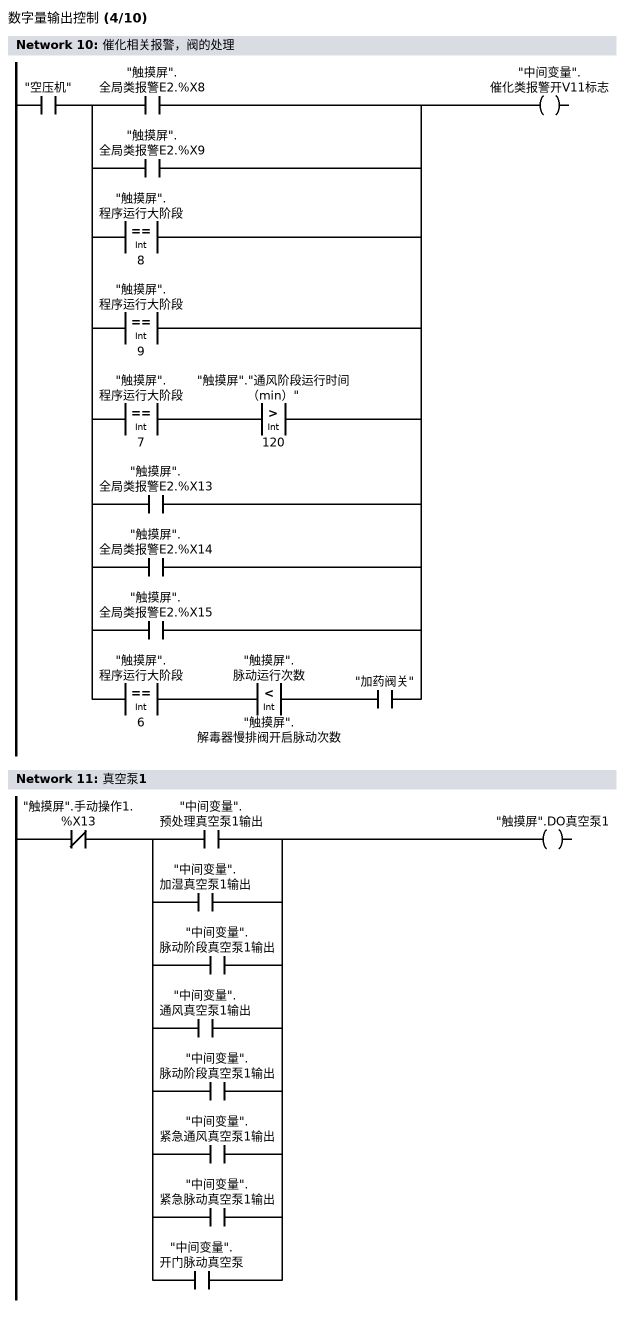
   RUNG wire#powerrail
      Contact( "空压机" )
      wire#w1
      Contact( "触摸屏".全局类报警E2.%X8 )
      wire#w2
      Coil( "中间变量".催化类报警开V11标志 )
   END_RUNG
   RUNG wire#w1
      Contact( "触摸屏".全局类报警E2.%X9 )
   END_RUNG wire#w2
   RUNG wire#w1
      { S7_Templates := "SrcType := Int" } EQ_Contact(in1 := "触摸屏".程序运行大阶段, in2 := 8)
   END_RUNG wire#w2
   RUNG wire#w1
      { S7_Templates := "SrcType := Int" } EQ_Contact(in1 := "触摸屏".程序运行大阶段, in2 := 9)
   END_RUNG wire#w2
   RUNG wire#w1
      { S7_Templates := "SrcType := Int" } EQ_Contact(in1 := "触摸屏".程序运行大阶段, in2 := 7)
      { S7_Templates := "SrcType := Int" } GT_Contact(in1 := "触摸屏"."通风阶段运行时间（min）", in2 := 120)
   END_RUNG wire#w2
   RUNG wire#w1
      Contact( "触摸屏".全局类报警E2.%X13 )
   END_RUNG wire#w2
   RUNG wire#w1
      Contact( "触摸屏".全局类报警E2.%X14 )
   END_RUNG wire#w2
   RUNG wire#w1
      Contact( "触摸屏".全局类报警E2.%X15 )
   END_RUNG wire#w2
   RUNG wire#w1
      { S7_Templates := "SrcType := Int" } EQ_Contact(in1 := "触摸屏".程序运行大阶段, in2 := 6)
      { S7_Templates := "SrcType := Int" } LT_Contact(in1 := "触摸屏".脉动运行次数, in2 := "触摸屏".解毒器慢排阀开启脉动次数)
      Contact( "加药阀关" )
   END_RUNG wire#w2
   // the same network as SCL:
   "中间变量".催化类报警开V11标志 := "空压机" AND ("触摸屏".全局类报警E2.%X8 OR "触摸屏".全局类报警E2.%X9 OR ("触摸屏".程序运行大阶段 = 8) OR ("触摸屏".程序运行大阶段 = 9) OR (("触摸屏".程序运行大阶段 = 7) AND ("触摸屏"."通风阶段运行时间（min）" > 120)) OR "触摸屏".全局类报警E2.%X13 OR "触摸屏".全局类报警E2.%X14 OR "触摸屏".全局类报警E2.%X15 OR (("触摸屏".程序运行大阶段 = 6) AND ("触摸屏".脉动运行次数 < "触摸屏".解毒器慢排阀开启脉动次数) AND "加药阀关"));
END_REGION

REGION Network 11: 真空泵1
   RUNG wire#powerrail
      I_Contact( "触摸屏".手动操作1.%X13 )
      wire#w1
      Contact( "中间变量".预处理真空泵1输出 )
      wire#w2
      Coil( "触摸屏".DO真空泵1 )
   END_RUNG
   RUNG wire#w1
      Contact( "中间变量".加湿真空泵1输出 )
   END_RUNG wire#w2
   RUNG wire#w1
      Contact( "中间变量".脉动阶段真空泵1输出 )
   END_RUNG wire#w2
   RUNG wire#w1
      Contact( "中间变量".通风真空泵1输出 )
   END_RUNG wire#w2
   RUNG wire#w1
      Contact( "中间变量".脉动阶段真空泵1输出 )
   END_RUNG wire#w2
   RUNG wire#w1
      Contact( "中间变量".紧急通风真空泵1输出 )
   END_RUNG wire#w2
   RUNG wire#w1
      Contact( "中间变量".紧急脉动真空泵1输出 )
   END_RUNG wire#w2
   RUNG wire#w1
      Contact( "中间变量".开门脉动真空泵 )
   END_RUNG wire#w2
   // the same network as SCL:
   "触摸屏".DO真空泵1 := NOT "触摸屏".手动操作1.%X13 AND ("中间变量".预处理真空泵1输出 OR "中间变量".加湿真空泵1输出 OR "中间变量".脉动阶段真空泵1输出 OR "中间变量".通风真空泵1输出 OR "中间变量".脉动阶段真空泵1输出 OR "中间变量".紧急通风真空泵1输出 OR "中间变量".紧急脉动真空泵1输出 OR "中间变量".开门脉动真空泵);
END_REGION

REGION Network 12: 真空泵2
END_REGION

REGION Network 13: 空压机
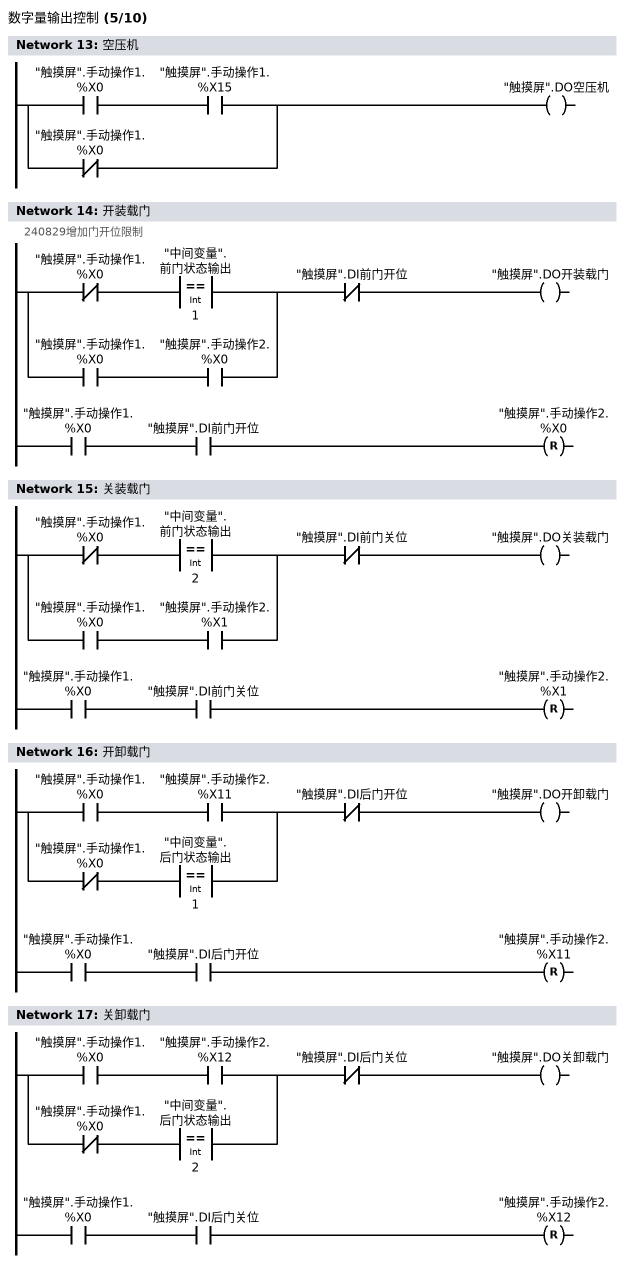
   RUNG wire#powerrail
      Contact( "触摸屏".手动操作1.%X0 )
      Contact( "触摸屏".手动操作1.%X15 )
      wire#w1
      Coil( "触摸屏".DO空压机 )
   END_RUNG
   RUNG wire#powerrail
      I_Contact( "触摸屏".手动操作1.%X0 )
   END_RUNG wire#w1
   // the same network as SCL:
   "触摸屏".DO空压机 := ("触摸屏".手动操作1.%X0 AND "触摸屏".手动操作1.%X15) OR NOT "触摸屏".手动操作1.%X0;
END_REGION

REGION Network 14: 开装载门
   // 240829增加门开位限制
   RUNG wire#powerrail
      I_Contact( "触摸屏".手动操作1.%X0 )
      { S7_Templates := "SrcType := Int" } EQ_Contact(in1 := "中间变量".前门状态输出, in2 := 1)
      wire#w1
      I_Contact( "触摸屏".DI前门开位 )
      Coil( "触摸屏".DO开装载门 )
   END_RUNG
   RUNG wire#powerrail
      Contact( "触摸屏".手动操作1.%X0 )
      Contact( "触摸屏".手动操作2.%X0 )
   END_RUNG wire#w1
   RUNG wire#powerrail
      Contact( "触摸屏".手动操作1.%X0 )
      Contact( "触摸屏".DI前门开位 )
      R_Coil( "触摸屏".手动操作2.%X0 )
   END_RUNG
   // the same network as SCL:
   "触摸屏".DO开装载门 := ((NOT "触摸屏".手动操作1.%X0 AND ("中间变量".前门状态输出 = 1)) OR ("触摸屏".手动操作1.%X0 AND "触摸屏".手动操作2.%X0)) AND NOT "触摸屏".DI前门开位;
   IF "触摸屏".手动操作1.%X0 AND "触摸屏".DI前门开位 THEN "触摸屏".手动操作2.%X0 := FALSE; END_IF;
END_REGION

REGION Network 15: 关装载门
   RUNG wire#powerrail
      I_Contact( "触摸屏".手动操作1.%X0 )
      { S7_Templates := "SrcType := Int" } EQ_Contact(in1 := "中间变量".前门状态输出, in2 := 2)
      wire#w1
      I_Contact( "触摸屏".DI前门关位 )
      Coil( "触摸屏".DO关装载门 )
   END_RUNG
   RUNG wire#powerrail
      Contact( "触摸屏".手动操作1.%X0 )
      Contact( "触摸屏".手动操作2.%X1 )
   END_RUNG wire#w1
   RUNG wire#powerrail
      Contact( "触摸屏".手动操作1.%X0 )
      Contact( "触摸屏".DI前门关位 )
      R_Coil( "触摸屏".手动操作2.%X1 )
   END_RUNG
   // the same network as SCL:
   "触摸屏".DO关装载门 := ((NOT "触摸屏".手动操作1.%X0 AND ("中间变量".前门状态输出 = 2)) OR ("触摸屏".手动操作1.%X0 AND "触摸屏".手动操作2.%X1)) AND NOT "触摸屏".DI前门关位;
   IF "触摸屏".手动操作1.%X0 AND "触摸屏".DI前门关位 THEN "触摸屏".手动操作2.%X1 := FALSE; END_IF;
END_REGION

REGION Network 16: 开卸载门
   RUNG wire#powerrail
      Contact( "触摸屏".手动操作1.%X0 )
      Contact( "触摸屏".手动操作2.%X11 )
      wire#w1
      I_Contact( "触摸屏".DI后门开位 )
      Coil( "触摸屏".DO开卸载门 )
   END_RUNG
   RUNG wire#powerrail
      I_Contact( "触摸屏".手动操作1.%X0 )
      { S7_Templates := "SrcType := Int" } EQ_Contact(in1 := "中间变量".后门状态输出, in2 := 1)
   END_RUNG wire#w1
   RUNG wire#powerrail
      Contact( "触摸屏".手动操作1.%X0 )
      Contact( "触摸屏".DI后门开位 )
      R_Coil( "触摸屏".手动操作2.%X11 )
   END_RUNG
   // the same network as SCL:
   "触摸屏".DO开卸载门 := (("触摸屏".手动操作1.%X0 AND "触摸屏".手动操作2.%X11) OR (NOT "触摸屏".手动操作1.%X0 AND ("中间变量".后门状态输出 = 1))) AND NOT "触摸屏".DI后门开位;
   IF "触摸屏".手动操作1.%X0 AND "触摸屏".DI后门开位 THEN "触摸屏".手动操作2.%X11 := FALSE; END_IF;
END_REGION

REGION Network 17: 关卸载门
   RUNG wire#powerrail
      Contact( "触摸屏".手动操作1.%X0 )
      Contact( "触摸屏".手动操作2.%X12 )
      wire#w1
      I_Contact( "触摸屏".DI后门关位 )
      Coil( "触摸屏".DO关卸载门 )
   END_RUNG
   RUNG wire#powerrail
      I_Contact( "触摸屏".手动操作1.%X0 )
      { S7_Templates := "SrcType := Int" } EQ_Contact(in1 := "中间变量".后门状态输出, in2 := 2)
   END_RUNG wire#w1
   RUNG wire#powerrail
      Contact( "触摸屏".手动操作1.%X0 )
      Contact( "触摸屏".DI后门关位 )
      R_Coil( "触摸屏".手动操作2.%X12 )
   END_RUNG
   // the same network as SCL:
   "触摸屏".DO关卸载门 := (("触摸屏".手动操作1.%X0 AND "触摸屏".手动操作2.%X12) OR (NOT "触摸屏".手动操作1.%X0 AND ("中间变量".后门状态输出 = 2))) AND NOT "触摸屏".DI后门关位;
   IF "触摸屏".手动操作1.%X0 AND "触摸屏".DI后门关位 THEN "触摸屏".手动操作2.%X12 := FALSE; END_IF;
END_REGION

REGION Network 18: 蜂鸣器FM
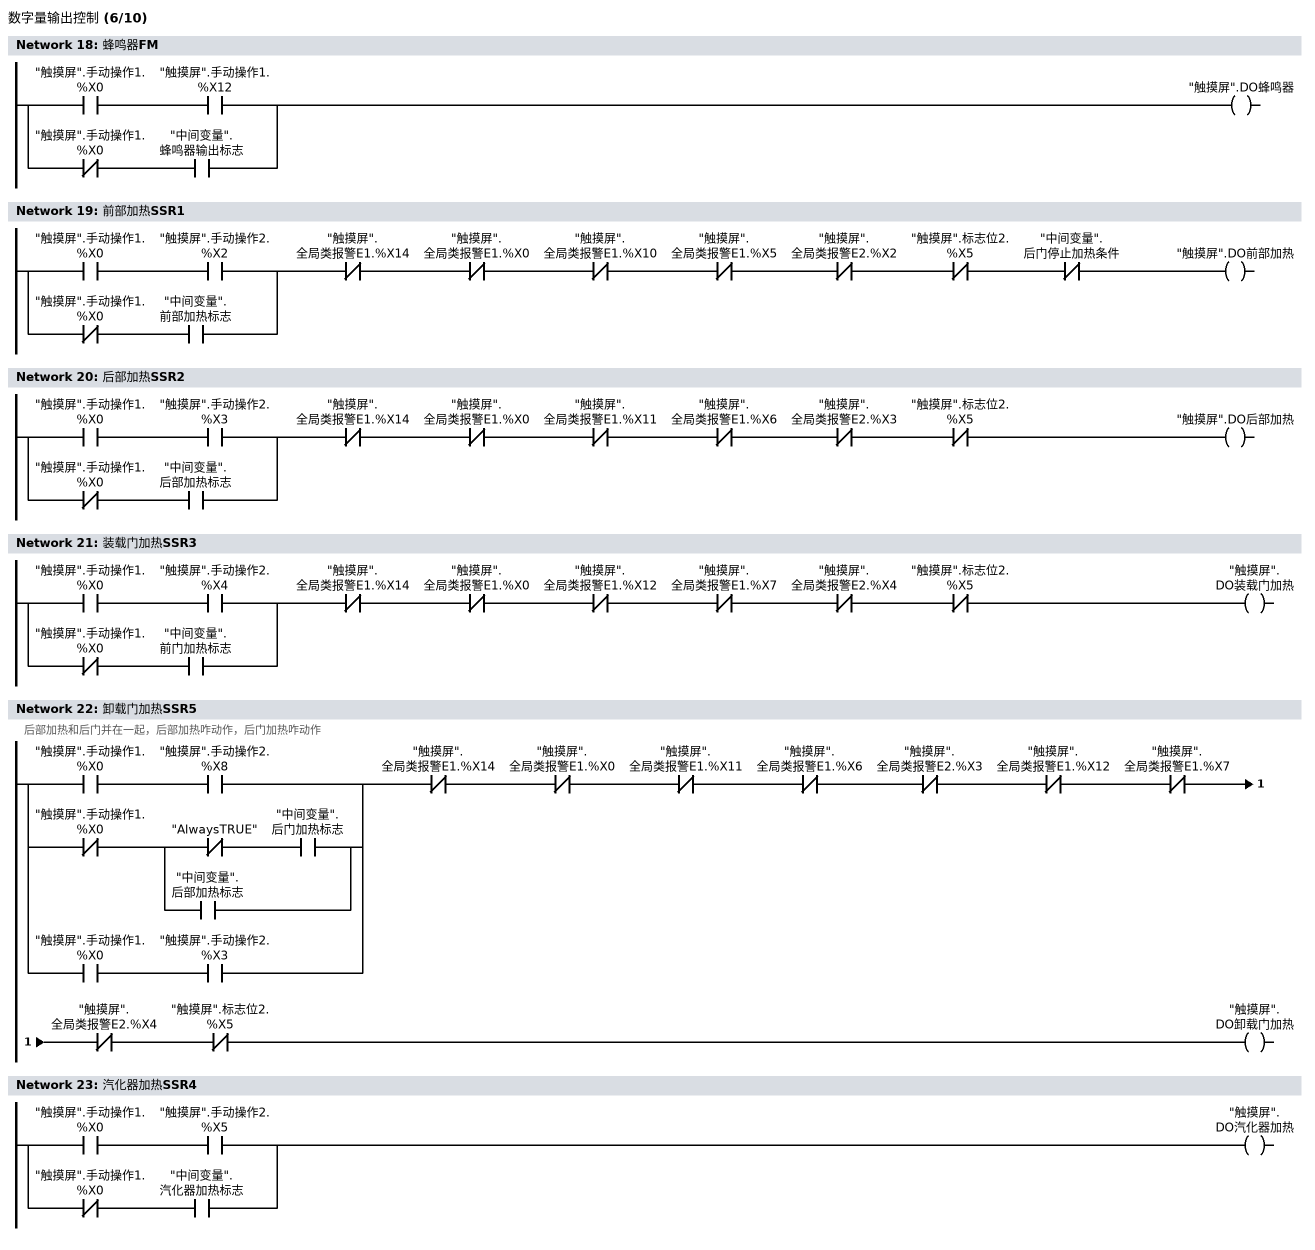
   RUNG wire#powerrail
      Contact( "触摸屏".手动操作1.%X0 )
      Contact( "触摸屏".手动操作1.%X12 )
      wire#w1
      Coil( "触摸屏".DO蜂鸣器 )
   END_RUNG
   RUNG wire#powerrail
      I_Contact( "触摸屏".手动操作1.%X0 )
      Contact( "中间变量".蜂鸣器输出标志 )
   END_RUNG wire#w1
   // the same network as SCL:
   "触摸屏".DO蜂鸣器 := ("触摸屏".手动操作1.%X0 AND "触摸屏".手动操作1.%X12) OR (NOT "触摸屏".手动操作1.%X0 AND "中间变量".蜂鸣器输出标志);
END_REGION

REGION Network 19: 前部加热SSR1
   RUNG wire#powerrail
      Contact( "触摸屏".手动操作1.%X0 )
      Contact( "触摸屏".手动操作2.%X2 )
      wire#w1
      I_Contact( "触摸屏".全局类报警E1.%X14 )
      I_Contact( "触摸屏".全局类报警E1.%X0 )
      I_Contact( "触摸屏".全局类报警E1.%X10 )
      I_Contact( "触摸屏".全局类报警E1.%X5 )
      I_Contact( "触摸屏".全局类报警E2.%X2 )
      I_Contact( "触摸屏".标志位2.%X5 )
      I_Contact( "中间变量".后门停止加热条件 )
      Coil( "触摸屏".DO前部加热 )
   END_RUNG
   RUNG wire#powerrail
      I_Contact( "触摸屏".手动操作1.%X0 )
      Contact( "中间变量".前部加热标志 )
   END_RUNG wire#w1
   // the same network as SCL:
   "触摸屏".DO前部加热 := (("触摸屏".手动操作1.%X0 AND "触摸屏".手动操作2.%X2) OR (NOT "触摸屏".手动操作1.%X0 AND "中间变量".前部加热标志)) AND NOT "触摸屏".全局类报警E1.%X14 AND NOT "触摸屏".全局类报警E1.%X0 AND NOT "触摸屏".全局类报警E1.%X10 AND NOT "触摸屏".全局类报警E1.%X5 AND NOT "触摸屏".全局类报警E2.%X2 AND NOT "触摸屏".标志位2.%X5 AND NOT "中间变量".后门停止加热条件;
END_REGION

REGION Network 20: 后部加热SSR2
   RUNG wire#powerrail
      Contact( "触摸屏".手动操作1.%X0 )
      Contact( "触摸屏".手动操作2.%X3 )
      wire#w1
      I_Contact( "触摸屏".全局类报警E1.%X14 )
      I_Contact( "触摸屏".全局类报警E1.%X0 )
      I_Contact( "触摸屏".全局类报警E1.%X11 )
      I_Contact( "触摸屏".全局类报警E1.%X6 )
      I_Contact( "触摸屏".全局类报警E2.%X3 )
      I_Contact( "触摸屏".标志位2.%X5 )
      Coil( "触摸屏".DO后部加热 )
   END_RUNG
   RUNG wire#powerrail
      I_Contact( "触摸屏".手动操作1.%X0 )
      Contact( "中间变量".后部加热标志 )
   END_RUNG wire#w1
   // the same network as SCL:
   "触摸屏".DO后部加热 := (("触摸屏".手动操作1.%X0 AND "触摸屏".手动操作2.%X3) OR (NOT "触摸屏".手动操作1.%X0 AND "中间变量".后部加热标志)) AND NOT "触摸屏".全局类报警E1.%X14 AND NOT "触摸屏".全局类报警E1.%X0 AND NOT "触摸屏".全局类报警E1.%X11 AND NOT "触摸屏".全局类报警E1.%X6 AND NOT "触摸屏".全局类报警E2.%X3 AND NOT "触摸屏".标志位2.%X5;
END_REGION

REGION Network 21: 装载门加热SSR3
   RUNG wire#powerrail
      Contact( "触摸屏".手动操作1.%X0 )
      Contact( "触摸屏".手动操作2.%X4 )
      wire#w1
      I_Contact( "触摸屏".全局类报警E1.%X14 )
      I_Contact( "触摸屏".全局类报警E1.%X0 )
      I_Contact( "触摸屏".全局类报警E1.%X12 )
      I_Contact( "触摸屏".全局类报警E1.%X7 )
      I_Contact( "触摸屏".全局类报警E2.%X4 )
      I_Contact( "触摸屏".标志位2.%X5 )
      Coil( "触摸屏".DO装载门加热 )
   END_RUNG
   RUNG wire#powerrail
      I_Contact( "触摸屏".手动操作1.%X0 )
      Contact( "中间变量".前门加热标志 )
   END_RUNG wire#w1
   // the same network as SCL:
   "触摸屏".DO装载门加热 := (("触摸屏".手动操作1.%X0 AND "触摸屏".手动操作2.%X4) OR (NOT "触摸屏".手动操作1.%X0 AND "中间变量".前门加热标志)) AND NOT "触摸屏".全局类报警E1.%X14 AND NOT "触摸屏".全局类报警E1.%X0 AND NOT "触摸屏".全局类报警E1.%X12 AND NOT "触摸屏".全局类报警E1.%X7 AND NOT "触摸屏".全局类报警E2.%X4 AND NOT "触摸屏".标志位2.%X5;
END_REGION

REGION Network 22: 卸载门加热SSR5
   // 后部加热和后门并在一起，后部加热咋动作，后门加热咋动作
   RUNG wire#powerrail
      Contact( "触摸屏".手动操作1.%X0 )
      Contact( "触摸屏".手动操作2.%X8 )
      wire#w1
      I_Contact( "触摸屏".全局类报警E1.%X14 )
      I_Contact( "触摸屏".全局类报警E1.%X0 )
      I_Contact( "触摸屏".全局类报警E1.%X11 )
      I_Contact( "触摸屏".全局类报警E1.%X6 )
      I_Contact( "触摸屏".全局类报警E2.%X3 )
      I_Contact( "触摸屏".全局类报警E1.%X12 )
      I_Contact( "触摸屏".全局类报警E1.%X7 )
      I_Contact( "触摸屏".全局类报警E2.%X4 )
      I_Contact( "触摸屏".标志位2.%X5 )
      Coil( "触摸屏".DO卸载门加热 )
   END_RUNG
   RUNG wire#powerrail
      I_Contact( "触摸屏".手动操作1.%X0 )
      wire#w2
      I_Contact( "AlwaysTRUE" )
      Contact( "中间变量".后门加热标志 )
   END_RUNG wire#w1
   RUNG wire#w2
      Contact( "中间变量".后部加热标志 )
   END_RUNG wire#w1
   RUNG wire#powerrail
      Contact( "触摸屏".手动操作1.%X0 )
      Contact( "触摸屏".手动操作2.%X3 )
   END_RUNG wire#w1
   // the same network as SCL:
   "触摸屏".DO卸载门加热 := (("触摸屏".手动操作1.%X0 AND "触摸屏".手动操作2.%X8) OR (NOT "触摸屏".手动操作1.%X0 AND ((NOT "AlwaysTRUE" AND "中间变量".后门加热标志) OR "中间变量".后部加热标志)) OR ("触摸屏".手动操作1.%X0 AND "触摸屏".手动操作2.%X3)) AND NOT "触摸屏".全局类报警E1.%X14 AND NOT "触摸屏".全局类报警E1.%X0 AND NOT "触摸屏".全局类报警E1.%X11 AND NOT "触摸屏".全局类报警E1.%X6 AND NOT "触摸屏".全局类报警E2.%X3 AND NOT "触摸屏".全局类报警E1.%X12 AND NOT "触摸屏".全局类报警E1.%X7 AND NOT "触摸屏".全局类报警E2.%X4 AND NOT "触摸屏".标志位2.%X5;
END_REGION

REGION Network 23: 汽化器加热SSR4
   RUNG wire#powerrail
      Contact( "触摸屏".手动操作1.%X0 )
      Contact( "触摸屏".手动操作2.%X5 )
      wire#w1
      Coil( "触摸屏".DO汽化器加热 )
   END_RUNG
   RUNG wire#powerrail
      I_Contact( "触摸屏".手动操作1.%X0 )
      Contact( "中间变量".汽化器加热标志 )
   END_RUNG wire#w1
   // the same network as SCL:
   "触摸屏".DO汽化器加热 := ("触摸屏".手动操作1.%X0 AND "触摸屏".手动操作2.%X5) OR (NOT "触摸屏".手动操作1.%X0 AND "中间变量".汽化器加热标志);
END_REGION

REGION Network 24: 催化加热1
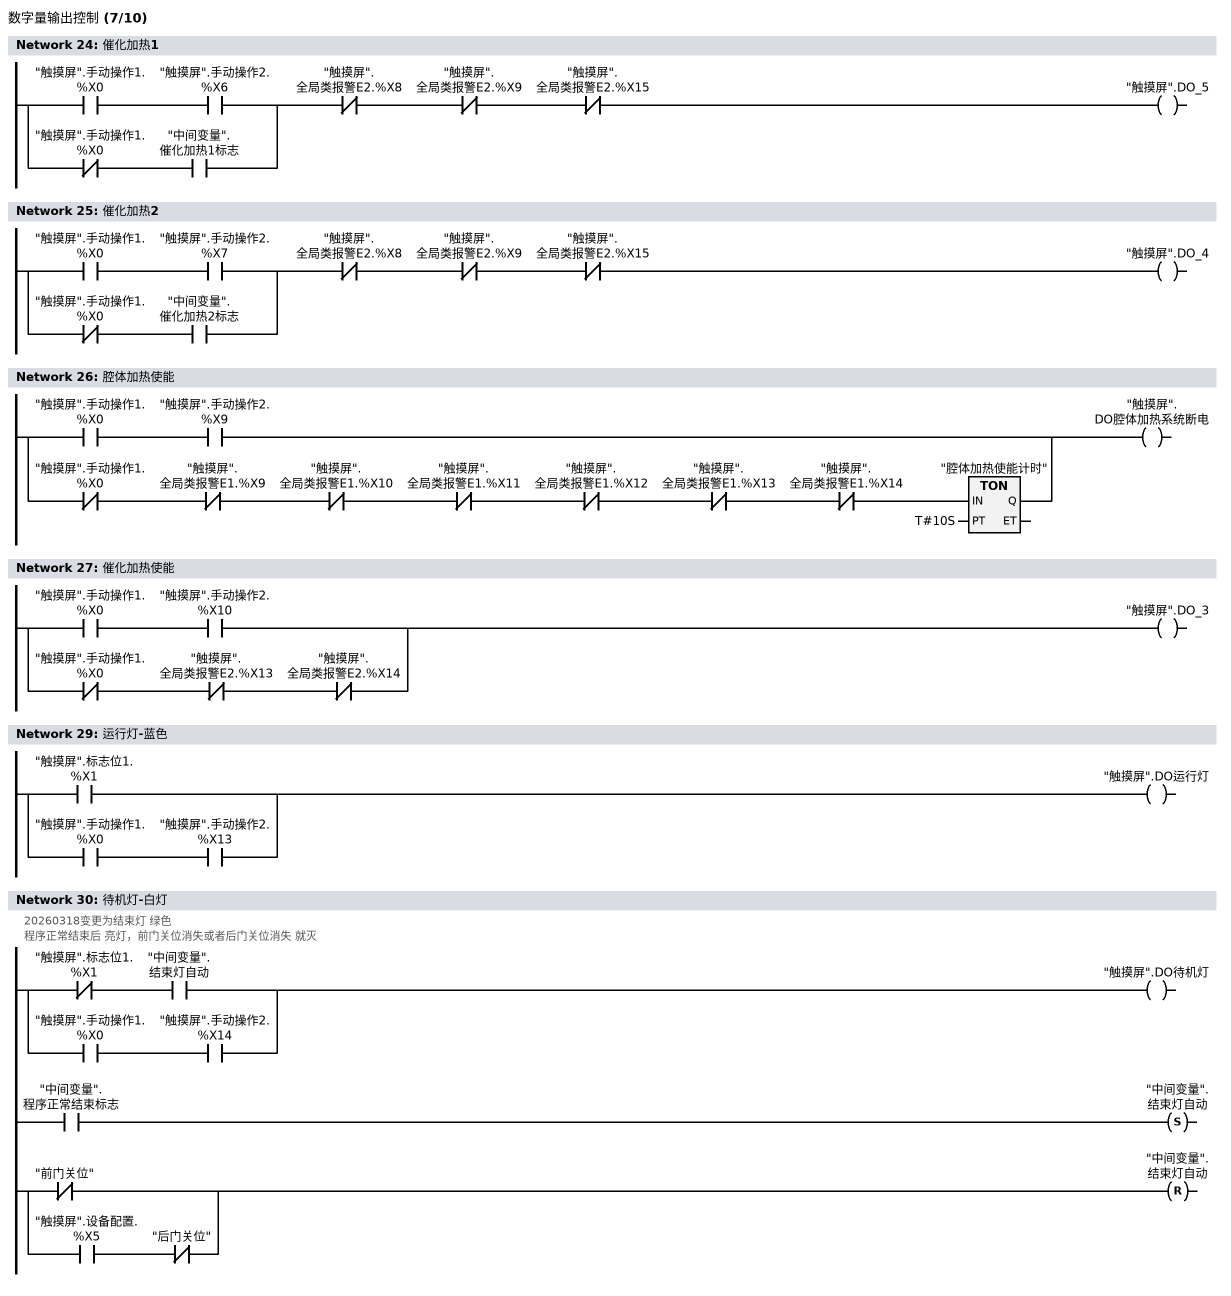
   RUNG wire#powerrail
      Contact( "触摸屏".手动操作1.%X0 )
      Contact( "触摸屏".手动操作2.%X6 )
      wire#w1
      I_Contact( "触摸屏".全局类报警E2.%X8 )
      I_Contact( "触摸屏".全局类报警E2.%X9 )
      I_Contact( "触摸屏".全局类报警E2.%X15 )
      Coil( "触摸屏".DO_5 )
   END_RUNG
   RUNG wire#powerrail
      I_Contact( "触摸屏".手动操作1.%X0 )
      Contact( "中间变量".催化加热1标志 )
   END_RUNG wire#w1
   // the same network as SCL:
   "触摸屏".DO_5 := (("触摸屏".手动操作1.%X0 AND "触摸屏".手动操作2.%X6) OR (NOT "触摸屏".手动操作1.%X0 AND "中间变量".催化加热1标志)) AND NOT "触摸屏".全局类报警E2.%X8 AND NOT "触摸屏".全局类报警E2.%X9 AND NOT "触摸屏".全局类报警E2.%X15;
END_REGION

REGION Network 25: 催化加热2
   RUNG wire#powerrail
      Contact( "触摸屏".手动操作1.%X0 )
      Contact( "触摸屏".手动操作2.%X7 )
      wire#w1
      I_Contact( "触摸屏".全局类报警E2.%X8 )
      I_Contact( "触摸屏".全局类报警E2.%X9 )
      I_Contact( "触摸屏".全局类报警E2.%X15 )
      Coil( "触摸屏".DO_4 )
   END_RUNG
   RUNG wire#powerrail
      I_Contact( "触摸屏".手动操作1.%X0 )
      Contact( "中间变量".催化加热2标志 )
   END_RUNG wire#w1
   // the same network as SCL:
   "触摸屏".DO_4 := (("触摸屏".手动操作1.%X0 AND "触摸屏".手动操作2.%X7) OR (NOT "触摸屏".手动操作1.%X0 AND "中间变量".催化加热2标志)) AND NOT "触摸屏".全局类报警E2.%X8 AND NOT "触摸屏".全局类报警E2.%X9 AND NOT "触摸屏".全局类报警E2.%X15;
END_REGION

REGION Network 26: 腔体加热使能
   "腔体加热使能计时".TON(IN := NOT "触摸屏".手动操作1.%X0 AND NOT "触摸屏".全局类报警E1.%X9 AND NOT "触摸屏".全局类报警E1.%X10 AND NOT "触摸屏".全局类报警E1.%X11 AND NOT "触摸屏".全局类报警E1.%X12 AND NOT "触摸屏".全局类报警E1.%X13 AND NOT "触摸屏".全局类报警E1.%X14,
                  PT := T#10S);
   "触摸屏".DO腔体加热系统断电 := ("触摸屏".手动操作1.%X0 AND "触摸屏".手动操作2.%X9) OR "腔体加热使能计时".Q;
END_REGION

REGION Network 27: 催化加热使能
   RUNG wire#powerrail
      Contact( "触摸屏".手动操作1.%X0 )
      Contact( "触摸屏".手动操作2.%X10 )
      wire#w1
      Coil( "触摸屏".DO_3 )
   END_RUNG
   RUNG wire#powerrail
      I_Contact( "触摸屏".手动操作1.%X0 )
      I_Contact( "触摸屏".全局类报警E2.%X13 )
      I_Contact( "触摸屏".全局类报警E2.%X14 )
   END_RUNG wire#w1
   // the same network as SCL:
   "触摸屏".DO_3 := ("触摸屏".手动操作1.%X0 AND "触摸屏".手动操作2.%X10) OR (NOT "触摸屏".手动操作1.%X0 AND NOT "触摸屏".全局类报警E2.%X13 AND NOT "触摸屏".全局类报警E2.%X14);
END_REGION

REGION Network 28: 脱扣器
END_REGION

REGION Network 29: 运行灯-蓝色
   RUNG wire#powerrail
      Contact( "触摸屏".标志位1.%X1 )
      wire#w1
      Coil( "触摸屏".DO运行灯 )
   END_RUNG
   RUNG wire#powerrail
      Contact( "触摸屏".手动操作1.%X0 )
      Contact( "触摸屏".手动操作2.%X13 )
   END_RUNG wire#w1
   // the same network as SCL:
   "触摸屏".DO运行灯 := "触摸屏".标志位1.%X1 OR ("触摸屏".手动操作1.%X0 AND "触摸屏".手动操作2.%X13);
END_REGION

REGION Network 30: 待机灯-白灯
   // 20260318变更为结束灯 绿色
   // 程序正常结束后 亮灯，前门关位消失或者后门关位消失 就灭
   RUNG wire#powerrail
      I_Contact( "触摸屏".标志位1.%X1 )
      Contact( "中间变量".结束灯自动 )
      wire#w1
      Coil( "触摸屏".DO待机灯 )
   END_RUNG
   RUNG wire#powerrail
      Contact( "触摸屏".手动操作1.%X0 )
      Contact( "触摸屏".手动操作2.%X14 )
   END_RUNG wire#w1
   RUNG wire#powerrail
      Contact( "中间变量".程序正常结束标志 )
      S_Coil( "中间变量".结束灯自动 )
   END_RUNG
   RUNG wire#powerrail
      I_Contact( "前门关位" )
      wire#w2
      R_Coil( "中间变量".结束灯自动 )
   END_RUNG
   RUNG wire#powerrail
      Contact( "触摸屏".设备配置.%X5 )
      I_Contact( "后门关位" )
   END_RUNG wire#w2
   // the same network as SCL:
   "触摸屏".DO待机灯 := (NOT "触摸屏".标志位1.%X1 AND "中间变量".结束灯自动) OR ("触摸屏".手动操作1.%X0 AND "触摸屏".手动操作2.%X14);
   IF "中间变量".程序正常结束标志 THEN "中间变量".结束灯自动 := TRUE; END_IF;
   IF NOT "前门关位" OR ("触摸屏".设备配置.%X5 AND NOT "后门关位") THEN "中间变量".结束灯自动 := FALSE; END_IF;
END_REGION

REGION Network 31: 报警灯-红灯
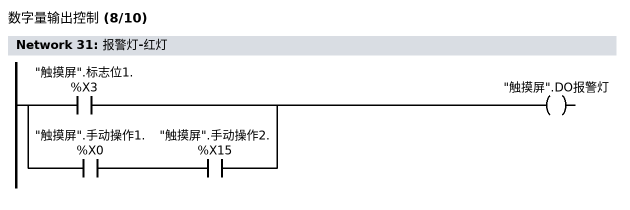
   RUNG wire#powerrail
      Contact( "触摸屏".标志位1.%X3 )
      wire#w1
      Coil( "触摸屏".DO报警灯 )
   END_RUNG
   RUNG wire#powerrail
      Contact( "触摸屏".手动操作1.%X0 )
      Contact( "触摸屏".手动操作2.%X15 )
   END_RUNG wire#w1
   // the same network as SCL:
   "触摸屏".DO报警灯 := "触摸屏".标志位1.%X3 OR ("触摸屏".手动操作1.%X0 AND "触摸屏".手动操作2.%X15);
END_REGION

REGION Network 32: 数字量输出信号全部转到DO输出映像区
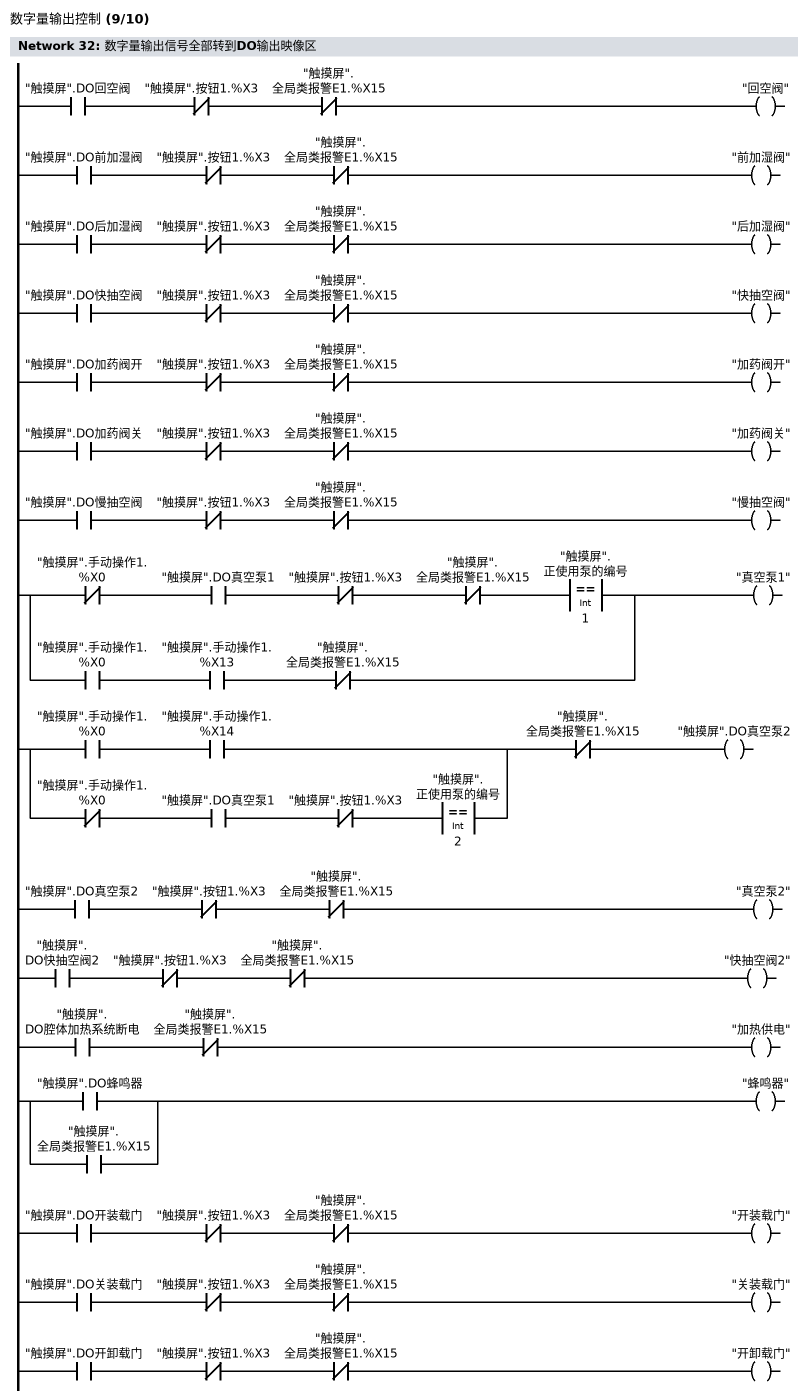
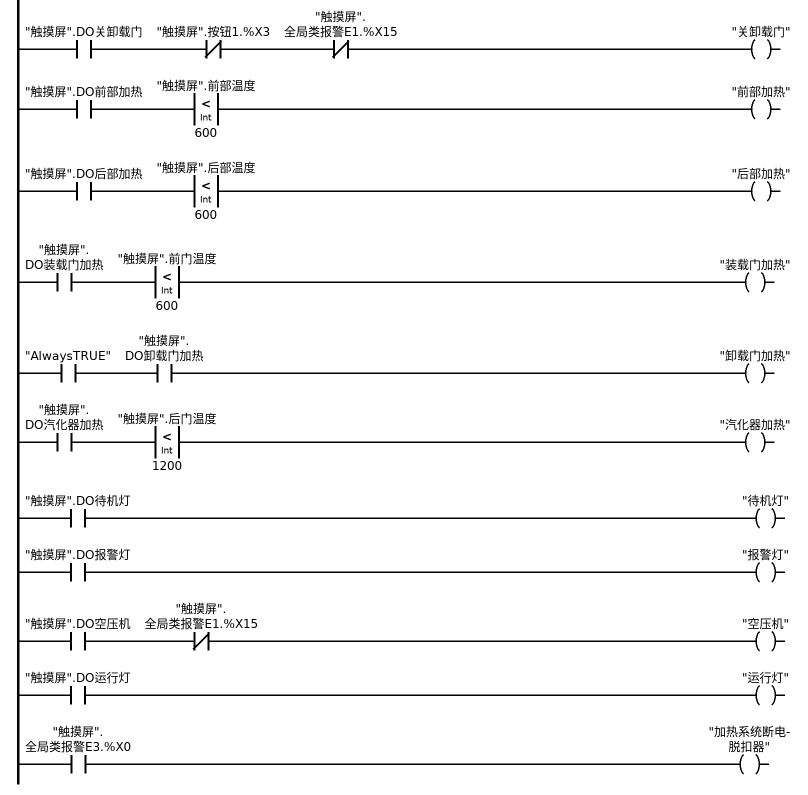
   RUNG wire#powerrail
      Contact( "触摸屏".DO回空阀 )
      I_Contact( "触摸屏".按钮1.%X3 )
      I_Contact( "触摸屏".全局类报警E1.%X15 )
      Coil( "回空阀" )
   END_RUNG
   RUNG wire#powerrail
      Contact( "触摸屏".DO前加湿阀 )
      I_Contact( "触摸屏".按钮1.%X3 )
      I_Contact( "触摸屏".全局类报警E1.%X15 )
      Coil( "前加湿阀" )
   END_RUNG
   RUNG wire#powerrail
      Contact( "触摸屏".DO后加湿阀 )
      I_Contact( "触摸屏".按钮1.%X3 )
      I_Contact( "触摸屏".全局类报警E1.%X15 )
      Coil( "后加湿阀" )
   END_RUNG
   RUNG wire#powerrail
      Contact( "触摸屏".DO快抽空阀 )
      I_Contact( "触摸屏".按钮1.%X3 )
      I_Contact( "触摸屏".全局类报警E1.%X15 )
      Coil( "快抽空阀" )
   END_RUNG
   RUNG wire#powerrail
      Contact( "触摸屏".DO加药阀开 )
      I_Contact( "触摸屏".按钮1.%X3 )
      I_Contact( "触摸屏".全局类报警E1.%X15 )
      Coil( "加药阀开" )
   END_RUNG
   RUNG wire#powerrail
      Contact( "触摸屏".DO加药阀关 )
      I_Contact( "触摸屏".按钮1.%X3 )
      I_Contact( "触摸屏".全局类报警E1.%X15 )
      Coil( "加药阀关" )
   END_RUNG
   RUNG wire#powerrail
      Contact( "触摸屏".DO慢抽空阀 )
      I_Contact( "触摸屏".按钮1.%X3 )
      I_Contact( "触摸屏".全局类报警E1.%X15 )
      Coil( "慢抽空阀" )
   END_RUNG
   RUNG wire#powerrail
      I_Contact( "触摸屏".手动操作1.%X0 )
      Contact( "触摸屏".DO真空泵1 )
      I_Contact( "触摸屏".按钮1.%X3 )
      I_Contact( "触摸屏".全局类报警E1.%X15 )
      { S7_Templates := "SrcType := Int" } EQ_Contact(in1 := "触摸屏".正使用泵的编号, in2 := 1)
      wire#w1
      Coil( "真空泵1" )
   END_RUNG
   RUNG wire#powerrail
      Contact( "触摸屏".手动操作1.%X0 )
      Contact( "触摸屏".手动操作1.%X13 )
      I_Contact( "触摸屏".全局类报警E1.%X15 )
   END_RUNG wire#w1
   RUNG wire#powerrail
      Contact( "触摸屏".手动操作1.%X0 )
      Contact( "触摸屏".手动操作1.%X14 )
      wire#w2
      I_Contact( "触摸屏".全局类报警E1.%X15 )
      Coil( "触摸屏".DO真空泵2 )
   END_RUNG
   RUNG wire#powerrail
      I_Contact( "触摸屏".手动操作1.%X0 )
      Contact( "触摸屏".DO真空泵1 )
      I_Contact( "触摸屏".按钮1.%X3 )
      { S7_Templates := "SrcType := Int" } EQ_Contact(in1 := "触摸屏".正使用泵的编号, in2 := 2)
   END_RUNG wire#w2
   RUNG wire#powerrail
      Contact( "触摸屏".DO真空泵2 )
      I_Contact( "触摸屏".按钮1.%X3 )
      I_Contact( "触摸屏".全局类报警E1.%X15 )
      Coil( "真空泵2" )
   END_RUNG
   RUNG wire#powerrail
      Contact( "触摸屏".DO快抽空阀2 )
      I_Contact( "触摸屏".按钮1.%X3 )
      I_Contact( "触摸屏".全局类报警E1.%X15 )
      Coil( "快抽空阀2" )
   END_RUNG
   RUNG wire#powerrail
      Contact( "触摸屏".DO腔体加热系统断电 )
      I_Contact( "触摸屏".全局类报警E1.%X15 )
      Coil( "加热供电" )
   END_RUNG
   RUNG wire#powerrail
      Contact( "触摸屏".DO蜂鸣器 )
      wire#w3
      Coil( "蜂鸣器" )
   END_RUNG
   RUNG wire#powerrail
      Contact( "触摸屏".全局类报警E1.%X15 )
   END_RUNG wire#w3
   RUNG wire#powerrail
      Contact( "触摸屏".DO开装载门 )
      I_Contact( "触摸屏".按钮1.%X3 )
      I_Contact( "触摸屏".全局类报警E1.%X15 )
      Coil( "开装载门" )
   END_RUNG
   RUNG wire#powerrail
      Contact( "触摸屏".DO关装载门 )
      I_Contact( "触摸屏".按钮1.%X3 )
      I_Contact( "触摸屏".全局类报警E1.%X15 )
      Coil( "关装载门" )
   END_RUNG
   RUNG wire#powerrail
      Contact( "触摸屏".DO开卸载门 )
      I_Contact( "触摸屏".按钮1.%X3 )
      I_Contact( "触摸屏".全局类报警E1.%X15 )
      Coil( "开卸载门" )
   END_RUNG
   RUNG wire#powerrail
      Contact( "触摸屏".DO关卸载门 )
      I_Contact( "触摸屏".按钮1.%X3 )
      I_Contact( "触摸屏".全局类报警E1.%X15 )
      Coil( "关卸载门" )
   END_RUNG
   RUNG wire#powerrail
      Contact( "触摸屏".DO前部加热 )
      { S7_Templates := "SrcType := Int" } LT_Contact(in1 := "触摸屏".前部温度, in2 := 600)
      Coil( "前部加热" )
   END_RUNG
   RUNG wire#powerrail
      Contact( "触摸屏".DO后部加热 )
      { S7_Templates := "SrcType := Int" } LT_Contact(in1 := "触摸屏".后部温度, in2 := 600)
      Coil( "后部加热" )
   END_RUNG
   RUNG wire#powerrail
      Contact( "触摸屏".DO装载门加热 )
      { S7_Templates := "SrcType := Int" } LT_Contact(in1 := "触摸屏".前门温度, in2 := 600)
      Coil( "装载门加热" )
   END_RUNG
   RUNG wire#powerrail
      Contact( "AlwaysTRUE" )
      Contact( "触摸屏".DO卸载门加热 )
      Coil( "卸载门加热" )
   END_RUNG
   RUNG wire#powerrail
      Contact( "触摸屏".DO汽化器加热 )
      { S7_Templates := "SrcType := Int" } LT_Contact(in1 := "触摸屏".后门温度, in2 := 1200)
      Coil( "汽化器加热" )
   END_RUNG
   RUNG wire#powerrail
      Contact( "触摸屏".DO待机灯 )
      Coil( "待机灯" )
   END_RUNG
   RUNG wire#powerrail
      Contact( "触摸屏".DO报警灯 )
      Coil( "报警灯" )
   END_RUNG
   RUNG wire#powerrail
      Contact( "触摸屏".DO空压机 )
      I_Contact( "触摸屏".全局类报警E1.%X15 )
      Coil( "空压机" )
   END_RUNG
   RUNG wire#powerrail
      Contact( "触摸屏".DO运行灯 )
      Coil( "运行灯" )
   END_RUNG
   RUNG wire#powerrail
      Contact( "触摸屏".全局类报警E3.%X0 )
      Coil( "加热系统断电-脱扣器" )
   END_RUNG
   // the same network as SCL:
   "回空阀" := "触摸屏".DO回空阀 AND NOT "触摸屏".按钮1.%X3 AND NOT "触摸屏".全局类报警E1.%X15;
   "前加湿阀" := "触摸屏".DO前加湿阀 AND NOT "触摸屏".按钮1.%X3 AND NOT "触摸屏".全局类报警E1.%X15;
   "后加湿阀" := "触摸屏".DO后加湿阀 AND NOT "触摸屏".按钮1.%X3 AND NOT "触摸屏".全局类报警E1.%X15;
   "快抽空阀" := "触摸屏".DO快抽空阀 AND NOT "触摸屏".按钮1.%X3 AND NOT "触摸屏".全局类报警E1.%X15;
   "加药阀开" := "触摸屏".DO加药阀开 AND NOT "触摸屏".按钮1.%X3 AND NOT "触摸屏".全局类报警E1.%X15;
   "加药阀关" := "触摸屏".DO加药阀关 AND NOT "触摸屏".按钮1.%X3 AND NOT "触摸屏".全局类报警E1.%X15;
   "慢抽空阀" := "触摸屏".DO慢抽空阀 AND NOT "触摸屏".按钮1.%X3 AND NOT "触摸屏".全局类报警E1.%X15;
   "真空泵1" := (NOT "触摸屏".手动操作1.%X0 AND "触摸屏".DO真空泵1 AND NOT "触摸屏".按钮1.%X3 AND NOT "触摸屏".全局类报警E1.%X15 AND ("触摸屏".正使用泵的编号 = 1)) OR ("触摸屏".手动操作1.%X0 AND "触摸屏".手动操作1.%X13 AND NOT "触摸屏".全局类报警E1.%X15);
   "触摸屏".DO真空泵2 := (("触摸屏".手动操作1.%X0 AND "触摸屏".手动操作1.%X14) OR (NOT "触摸屏".手动操作1.%X0 AND "触摸屏".DO真空泵1 AND NOT "触摸屏".按钮1.%X3 AND ("触摸屏".正使用泵的编号 = 2))) AND NOT "触摸屏".全局类报警E1.%X15;
   "真空泵2" := "触摸屏".DO真空泵2 AND NOT "触摸屏".按钮1.%X3 AND NOT "触摸屏".全局类报警E1.%X15;
   "快抽空阀2" := "触摸屏".DO快抽空阀2 AND NOT "触摸屏".按钮1.%X3 AND NOT "触摸屏".全局类报警E1.%X15;
   "加热供电" := "触摸屏".DO腔体加热系统断电 AND NOT "触摸屏".全局类报警E1.%X15;
   "蜂鸣器" := "触摸屏".DO蜂鸣器 OR "触摸屏".全局类报警E1.%X15;
   "开装载门" := "触摸屏".DO开装载门 AND NOT "触摸屏".按钮1.%X3 AND NOT "触摸屏".全局类报警E1.%X15;
   "关装载门" := "触摸屏".DO关装载门 AND NOT "触摸屏".按钮1.%X3 AND NOT "触摸屏".全局类报警E1.%X15;
   "开卸载门" := "触摸屏".DO开卸载门 AND NOT "触摸屏".按钮1.%X3 AND NOT "触摸屏".全局类报警E1.%X15;
   "关卸载门" := "触摸屏".DO关卸载门 AND NOT "触摸屏".按钮1.%X3 AND NOT "触摸屏".全局类报警E1.%X15;
   "前部加热" := "触摸屏".DO前部加热 AND ("触摸屏".前部温度 < 600);
   "后部加热" := "触摸屏".DO后部加热 AND ("触摸屏".后部温度 < 600);
   "装载门加热" := "触摸屏".DO装载门加热 AND ("触摸屏".前门温度 < 600);
   "卸载门加热" := "AlwaysTRUE" AND "触摸屏".DO卸载门加热;
   "汽化器加热" := "触摸屏".DO汽化器加热 AND ("触摸屏".后门温度 < 1200);
   "待机灯" := "触摸屏".DO待机灯;
   "报警灯" := "触摸屏".DO报警灯;
   "空压机" := "触摸屏".DO空压机 AND NOT "触摸屏".全局类报警E1.%X15;
   "运行灯" := "触摸屏".DO运行灯;
   "加热系统断电-脱扣器" := "触摸屏".全局类报警E3.%X0;
END_REGION

REGION Network 33: 手动操作变量清零
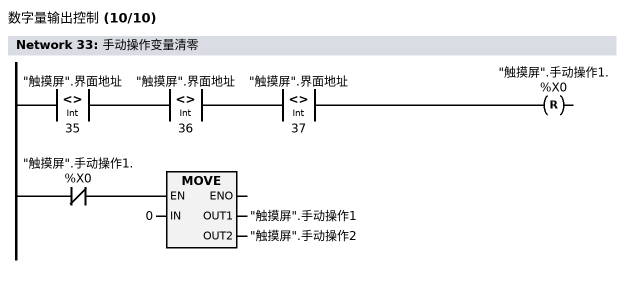
   RUNG wire#powerrail
      { S7_Templates := "SrcType := Int" } NE_Contact(in1 := "触摸屏".界面地址, in2 := 35)
      { S7_Templates := "SrcType := Int" } NE_Contact(in1 := "触摸屏".界面地址, in2 := 36)
      { S7_Templates := "SrcType := Int" } NE_Contact(in1 := "触摸屏".界面地址, in2 := 37)
      R_Coil( "触摸屏".手动操作1.%X0 )
   END_RUNG
   RUNG wire#powerrail
      I_Contact( "触摸屏".手动操作1.%X0 )
      Move(in := 0, out1 => "触摸屏".手动操作1, out2 => "触摸屏".手动操作2)
   END_RUNG
   // the same network as SCL:
   IF ("触摸屏".界面地址 <> 35) AND ("触摸屏".界面地址 <> 36) AND ("触摸屏".界面地址 <> 37) THEN "触摸屏".手动操作1.%X0 := FALSE; END_IF;
   IF NOT "触摸屏".手动操作1.%X0 THEN
       "触摸屏".手动操作1 := 0;
       "触摸屏".手动操作2 := 0;
   END_IF;
END_REGION
END_FUNCTION

// folder: 17页面控制

FUNCTION_BLOCK "页面跳转控制"   // FB20, LAD
{ S7_Optimized_Access := 'TRUE' }
VERSION : 0.1
   VAR RETAIN
      沿1 : Bool;
   END_VAR
   VAR
      沿2 : Bool;
   END_VAR
   VAR RETAIN
      新报警产生上升沿 : Bool;
      程序运行结束下降沿 : Bool;
      报警确认按钮沿 : Bool;
      程序异常运行结束下降沿 : Bool;
      泄露测试结束沿 : Bool;
   END_VAR
   VAR
      进入到预热选择页面沿 : Bool;
   END_VAR
   VAR_TEMP   // added for the SCL form of the ladder/FBD networks
      _w1 : Bool;
      _w2 : Bool;
      _w3 : Bool;
      _w4 : Bool;
      _w5 : Bool;
      _w6 : Bool;
   END_VAR
BEGIN

REGION Network 1: 本地大气压设置页面
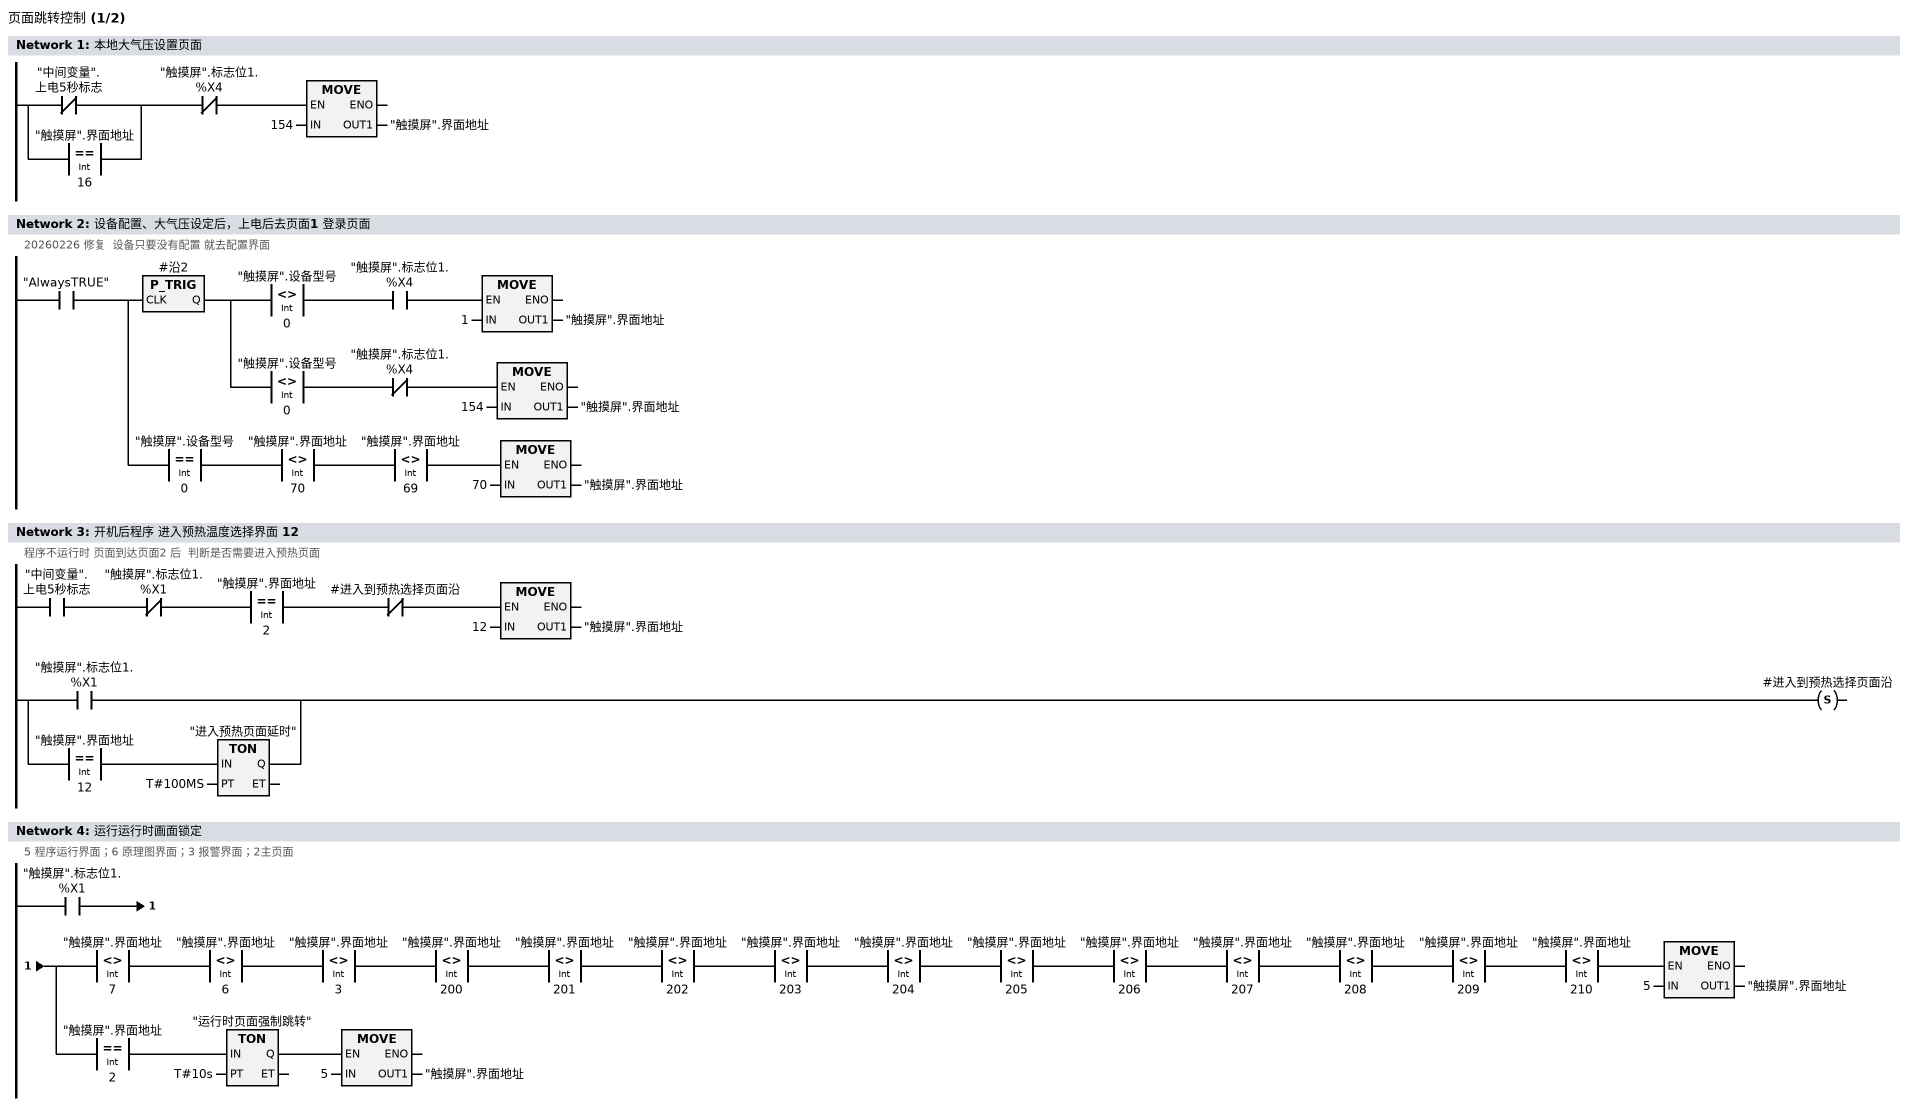
   RUNG wire#powerrail
      I_Contact( "中间变量".上电5秒标志 )
      wire#w1
      I_Contact( "触摸屏".标志位1.%X4 )
      Move(in := 154, out1 => "触摸屏".界面地址)
   END_RUNG
   RUNG wire#powerrail
      { S7_Templates := "SrcType := Int" } EQ_Contact(in1 := "触摸屏".界面地址, in2 := 16)
   END_RUNG wire#w1
   // the same network as SCL:
   IF (NOT "中间变量".上电5秒标志 OR ("触摸屏".界面地址 = 16)) AND NOT "触摸屏".标志位1.%X4 THEN "触摸屏".界面地址 := 154; END_IF;
END_REGION

REGION Network 2: 设备配置、大气压设定后，上电后去页面1 登录页面
   // 20260226 修复  设备只要没有配置 就去配置界面
   RUNG wire#powerrail
      Contact( "AlwaysTRUE" )
      wire#w1
      P_Trig( #沿2 )
      wire#w2
      { S7_Templates := "SrcType := Int" } NE_Contact(in1 := "触摸屏".设备型号, in2 := 0)
      Contact( "触摸屏".标志位1.%X4 )
      Move(in := 1, out1 => "触摸屏".界面地址)
   END_RUNG
   RUNG wire#w2
      { S7_Templates := "SrcType := Int" } NE_Contact(in1 := "触摸屏".设备型号, in2 := 0)
      I_Contact( "触摸屏".标志位1.%X4 )
      Move(in := 154, out1 => "触摸屏".界面地址)
   END_RUNG
   RUNG wire#w1
      { S7_Templates := "SrcType := Int" } EQ_Contact(in1 := "触摸屏".设备型号, in2 := 0)
      { S7_Templates := "SrcType := Int" } NE_Contact(in1 := "触摸屏".界面地址, in2 := 70)
      { S7_Templates := "SrcType := Int" } NE_Contact(in1 := "触摸屏".界面地址, in2 := 69)
      Move(in := 70, out1 => "触摸屏".界面地址)
   END_RUNG
   // the same network as SCL:
   #_w1 := "AlwaysTRUE" AND NOT #沿2;   // rising edge
   #沿2 := "AlwaysTRUE";
   IF #_w1 AND ("触摸屏".设备型号 <> 0) AND "触摸屏".标志位1.%X4 THEN "触摸屏".界面地址 := 1; END_IF;
   IF #_w1 AND ("触摸屏".设备型号 <> 0) AND NOT "触摸屏".标志位1.%X4 THEN "触摸屏".界面地址 := 154; END_IF;
   IF "AlwaysTRUE" AND ("触摸屏".设备型号 = 0) AND ("触摸屏".界面地址 <> 70) AND ("触摸屏".界面地址 <> 69) THEN
       "触摸屏".界面地址 := 70;
   END_IF;
END_REGION

REGION Network 3: 开机后程序 进入预热温度选择界面 12
   // 程序不运行时 页面到达页面2 后  判断是否需要进入预热页面
   IF "中间变量".上电5秒标志 AND NOT "触摸屏".标志位1.%X1 AND ("触摸屏".界面地址 = 2) AND NOT #进入到预热选择页面沿 THEN
       "触摸屏".界面地址 := 12;
   END_IF;
   "进入预热页面延时".TON(IN := "触摸屏".界面地址 = 12, PT := T#100MS);
   IF "触摸屏".标志位1.%X1 OR "进入预热页面延时".Q THEN #进入到预热选择页面沿 := TRUE; END_IF;
END_REGION

REGION Network 4: 运行运行时画面锁定
   // 5 程序运行界面；6 原理图界面；3 报警界面；2主页面
   IF "触摸屏".标志位1.%X1 AND ("触摸屏".界面地址 <> 7) AND ("触摸屏".界面地址 <> 6) AND ("触摸屏".界面地址 <> 3) AND ("触摸屏".界面地址 <> 200) AND ("触摸屏".界面地址 <> 201) AND ("触摸屏".界面地址 <> 202) AND ("触摸屏".界面地址 <> 203) AND ("触摸屏".界面地址 <> 204) AND ("触摸屏".界面地址 <> 205) AND ("触摸屏".界面地址 <> 206) AND ("触摸屏".界面地址 <> 207) AND ("触摸屏".界面地址 <> 208) AND ("触摸屏".界面地址 <> 209) AND ("触摸屏".界面地址 <> 210) THEN
       "触摸屏".界面地址 := 5;
   END_IF;
   "运行时页面强制跳转".TON(IN := "触摸屏".标志位1.%X1 AND ("触摸屏".界面地址 = 2), PT := T#10s);
   IF "运行时页面强制跳转".Q THEN "触摸屏".界面地址 := 5; END_IF;
END_REGION

REGION Network 5: 程序结束后点“主菜单”按钮页面跳转
   // 1.该按钮要做的事情有    催化剂过期报警       、页面跳转
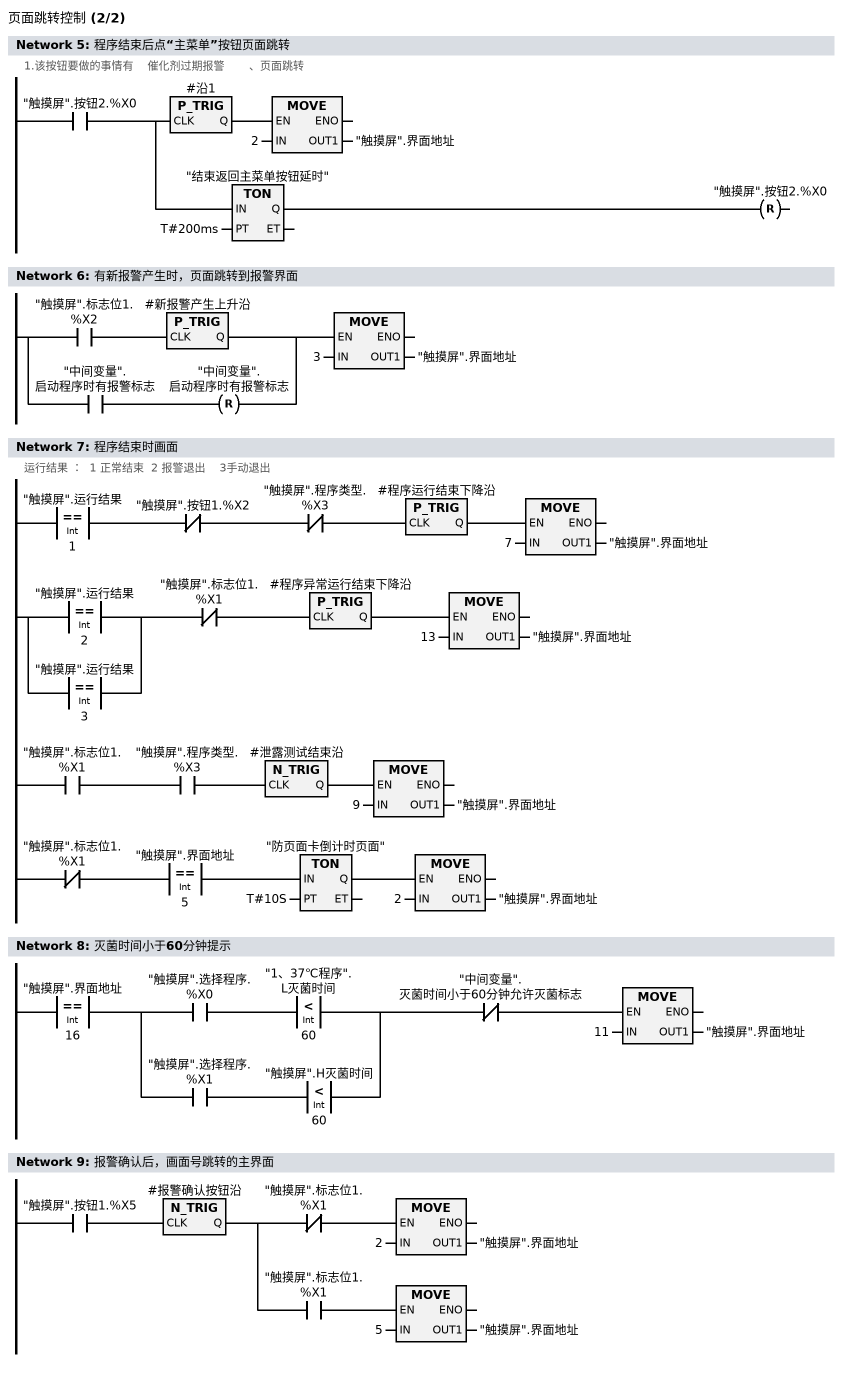
   #_w1 := "触摸屏".按钮2.%X0 AND NOT #沿1;   // rising edge
   #沿1 := "触摸屏".按钮2.%X0;
   IF #_w1 THEN "触摸屏".界面地址 := 2; END_IF;
   "结束返回主菜单按钮延时".TON(IN := "触摸屏".按钮2.%X0, PT := T#200ms);
   IF "结束返回主菜单按钮延时".Q THEN "触摸屏".按钮2.%X0 := FALSE; END_IF;
END_REGION

REGION Network 6: 有新报警产生时，页面跳转到报警界面
   RUNG wire#powerrail
      Contact( "触摸屏".标志位1.%X2 )
      P_Trig( #新报警产生上升沿 )
      wire#w1
      Move(in := 3, out1 => "触摸屏".界面地址)
   END_RUNG
   RUNG wire#powerrail
      Contact( "中间变量".启动程序时有报警标志 )
      R_Coil( "中间变量".启动程序时有报警标志 )
   END_RUNG wire#w1
   // the same network as SCL:
   #_w1 := "触摸屏".标志位1.%X2 AND NOT #新报警产生上升沿;   // rising edge
   #新报警产生上升沿 := "触摸屏".标志位1.%X2;
   #_w2 := "中间变量".启动程序时有报警标志;
   IF #_w2 THEN "中间变量".启动程序时有报警标志 := FALSE; END_IF;
   IF #_w1 OR #_w2 THEN "触摸屏".界面地址 := 3; END_IF;
END_REGION

REGION Network 7: 程序结束时画面
   // 运行结果 ：  1 正常结束  2 报警退出    3手动退出
   #_w1 := ("触摸屏".运行结果 = 1) AND NOT "触摸屏".按钮1.%X2 AND NOT "触摸屏".程序类型.%X3;
   #_w2 := #_w1 AND NOT #程序运行结束下降沿;   // rising edge
   #程序运行结束下降沿 := #_w1;
   IF #_w2 THEN "触摸屏".界面地址 := 7; END_IF;
   #_w3 := (("触摸屏".运行结果 = 2) OR ("触摸屏".运行结果 = 3)) AND NOT "触摸屏".标志位1.%X1;
   #_w4 := #_w3 AND NOT #程序异常运行结束下降沿;   // rising edge
   #程序异常运行结束下降沿 := #_w3;
   IF #_w4 THEN "触摸屏".界面地址 := 13; END_IF;
   #_w5 := "触摸屏".标志位1.%X1 AND "触摸屏".程序类型.%X3;
   #_w6 := NOT #_w5 AND #泄露测试结束沿;   // falling edge
   #泄露测试结束沿 := #_w5;
   IF #_w6 THEN "触摸屏".界面地址 := 9; END_IF;
   "防页面卡倒计时页面".TON(IN := NOT "触摸屏".标志位1.%X1 AND ("触摸屏".界面地址 = 5), PT := T#10S);
   IF "防页面卡倒计时页面".Q THEN "触摸屏".界面地址 := 2; END_IF;
END_REGION

REGION Network 8: 灭菌时间小于60分钟提示
   RUNG wire#powerrail
      { S7_Templates := "SrcType := Int" } EQ_Contact(in1 := "触摸屏".界面地址, in2 := 16)
      wire#w1
      Contact( "触摸屏".选择程序.%X0 )
      { S7_Templates := "SrcType := Int" } LT_Contact(in1 := "1、37℃程序".L灭菌时间, in2 := 60)
      wire#w2
      I_Contact( "中间变量".灭菌时间小于60分钟允许灭菌标志 )
      Move(in := 11, out1 => "触摸屏".界面地址)
   END_RUNG
   RUNG wire#w1
      Contact( "触摸屏".选择程序.%X1 )
      { S7_Templates := "SrcType := Int" } LT_Contact(in1 := "触摸屏".H灭菌时间, in2 := 60)
   END_RUNG wire#w2
   // the same network as SCL:
   IF ("触摸屏".界面地址 = 16) AND (("触摸屏".选择程序.%X0 AND ("1、37℃程序".L灭菌时间 < 60)) OR ("触摸屏".选择程序.%X1 AND ("触摸屏".H灭菌时间 < 60))) AND NOT "中间变量".灭菌时间小于60分钟允许灭菌标志 THEN
       "触摸屏".界面地址 := 11;
   END_IF;
END_REGION

REGION Network 9: 报警确认后，画面号跳转的主界面
   RUNG wire#powerrail
      Contact( "触摸屏".按钮1.%X5 )
      N_Trig( #报警确认按钮沿 )
      wire#w1
      I_Contact( "触摸屏".标志位1.%X1 )
      Move(in := 2, out1 => "触摸屏".界面地址)
   END_RUNG
   RUNG wire#w1
      Contact( "触摸屏".标志位1.%X1 )
      Move(in := 5, out1 => "触摸屏".界面地址)
   END_RUNG
   // the same network as SCL:
   #_w1 := NOT "触摸屏".按钮1.%X5 AND #报警确认按钮沿;   // falling edge
   #报警确认按钮沿 := "触摸屏".按钮1.%X5;
   IF #_w1 AND NOT "触摸屏".标志位1.%X1 THEN "触摸屏".界面地址 := 2; END_IF;
   IF #_w1 AND "触摸屏".标志位1.%X1 THEN "触摸屏".界面地址 := 5; END_IF;
END_REGION

REGION Network 10: 加水完成页面跳转
END_REGION
END_FUNCTION_BLOCK

// folder: 200尾气处理器

FUNCTION_BLOCK "尾气处理器处理"   // FB24, LAD
TITLE = 不要使用外边变量 保持程序块的独立性
{ S7_Optimized_Access := 'TRUE' }
VERSION : 0.1
   VAR_OUTPUT
      与REO通讯故障标志_1 : Bool;
   END_VAR
   VAR
      心跳沿1 : Bool;
      心跳沿2 : Bool;
      沿预留0 : Bool;
      沿预留1 : Bool;
      沿预留2 : Bool;
      沿预留3 : Bool;
      沿预留4 : Bool;
      沿预留5 : Bool;
      沿预留6 : Bool;
      沿预留7 : Bool;
      沿预留8 : Bool;
      沿预留9 : Bool;
      沿预留10 : Bool;
      沿预留11 : Bool;
      沿预留12 : Bool;
      沿预留13 : Bool;
      灭菌剩余时间 : Int;
      按钮延时复位 : TON_TIME;
      REO通讯故障延时 : TON_TIME;
      REO心跳缓存数据 : Int;
   END_VAR
   VAR_TEMP   // added for the SCL form of the ladder/FBD networks
      _w1 : Bool;
      _w2 : Bool;
   END_VAR
BEGIN

REGION Network 1: 与尾气处理器的通讯状态
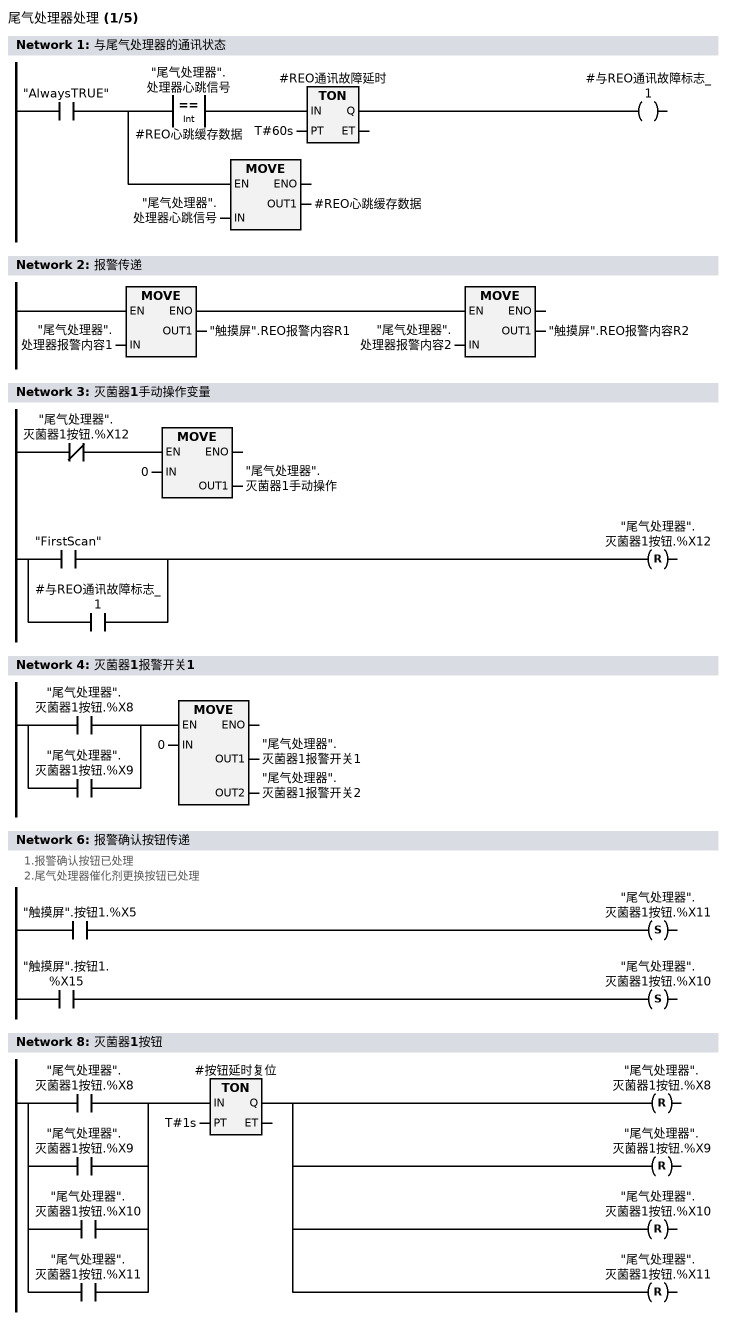
   #REO通讯故障延时(IN := "AlwaysTRUE" AND ("尾气处理器".处理器心跳信号 = #REO心跳缓存数据), PT := T#60s);   // TON
   #与REO通讯故障标志_1 := #REO通讯故障延时.Q;
   IF "AlwaysTRUE" THEN #REO心跳缓存数据 := "尾气处理器".处理器心跳信号; END_IF;
END_REGION

REGION Network 2: 报警传递
   RUNG wire#powerrail
      Move(in := "尾气处理器".处理器报警内容1, out1 => "触摸屏".REO报警内容R1)
      Move(in := "尾气处理器".处理器报警内容2, out1 => "触摸屏".REO报警内容R2)
   END_RUNG
   // the same network as SCL:
   "触摸屏".REO报警内容R1 := "尾气处理器".处理器报警内容1;
   "触摸屏".REO报警内容R2 := "尾气处理器".处理器报警内容2;
END_REGION

REGION Network 3: 灭菌器1手动操作变量
   RUNG wire#powerrail
      I_Contact( "尾气处理器".灭菌器1按钮.%X12 )
      Move(in := 0, out1 => "尾气处理器".灭菌器1手动操作)
   END_RUNG
   RUNG wire#powerrail
      Contact( "FirstScan" )
      wire#w1
      R_Coil( "尾气处理器".灭菌器1按钮.%X12 )
   END_RUNG
   RUNG wire#powerrail
      Contact( #与REO通讯故障标志_1 )
   END_RUNG wire#w1
   // the same network as SCL:
   IF NOT "尾气处理器".灭菌器1按钮.%X12 THEN "尾气处理器".灭菌器1手动操作 := 0; END_IF;
   IF "FirstScan" OR #与REO通讯故障标志_1 THEN "尾气处理器".灭菌器1按钮.%X12 := FALSE; END_IF;
END_REGION

REGION Network 4: 灭菌器1报警开关1
   RUNG wire#powerrail
      Contact( "尾气处理器".灭菌器1按钮.%X8 )
      wire#w1
      Move(in := 0, out1 => "尾气处理器".灭菌器1报警开关1, out2 => "尾气处理器".灭菌器1报警开关2)
   END_RUNG
   RUNG wire#powerrail
      Contact( "尾气处理器".灭菌器1按钮.%X9 )
   END_RUNG wire#w1
   // the same network as SCL:
   IF "尾气处理器".灭菌器1按钮.%X8 OR "尾气处理器".灭菌器1按钮.%X9 THEN
       "尾气处理器".灭菌器1报警开关1 := 0;
       "尾气处理器".灭菌器1报警开关2 := 0;
   END_IF;
END_REGION

REGION Network 5: 灭菌器1报警开关2
END_REGION

REGION Network 6: 报警确认按钮传递
   // 1.报警确认按钮已处理
   // 2.尾气处理器催化剂更换按钮已处理
   RUNG wire#powerrail
      Contact( "触摸屏".按钮1.%X5 )
      S_Coil( "尾气处理器".灭菌器1按钮.%X11 )
   END_RUNG
   RUNG wire#powerrail
      Contact( "触摸屏".按钮1.%X15 )
      S_Coil( "尾气处理器".灭菌器1按钮.%X10 )
   END_RUNG
   // the same network as SCL:
   IF "触摸屏".按钮1.%X5 THEN "尾气处理器".灭菌器1按钮.%X11 := TRUE; END_IF;
   IF "触摸屏".按钮1.%X15 THEN "尾气处理器".灭菌器1按钮.%X10 := TRUE; END_IF;
END_REGION

REGION Network 8: 灭菌器1按钮
   #按钮延时复位(IN := "尾气处理器".灭菌器1按钮.%X8 OR "尾气处理器".灭菌器1按钮.%X9 OR "尾气处理器".灭菌器1按钮.%X10 OR "尾气处理器".灭菌器1按钮.%X11,   // TON
           PT := T#1s);
   IF #按钮延时复位.Q THEN
       "尾气处理器".灭菌器1按钮.%X8 := FALSE;
       "尾气处理器".灭菌器1按钮.%X9 := FALSE;
       "尾气处理器".灭菌器1按钮.%X10 := FALSE;
       "尾气处理器".灭菌器1按钮.%X11 := FALSE;
   END_IF;
END_REGION

REGION Network 9: 灭菌器1大阶段
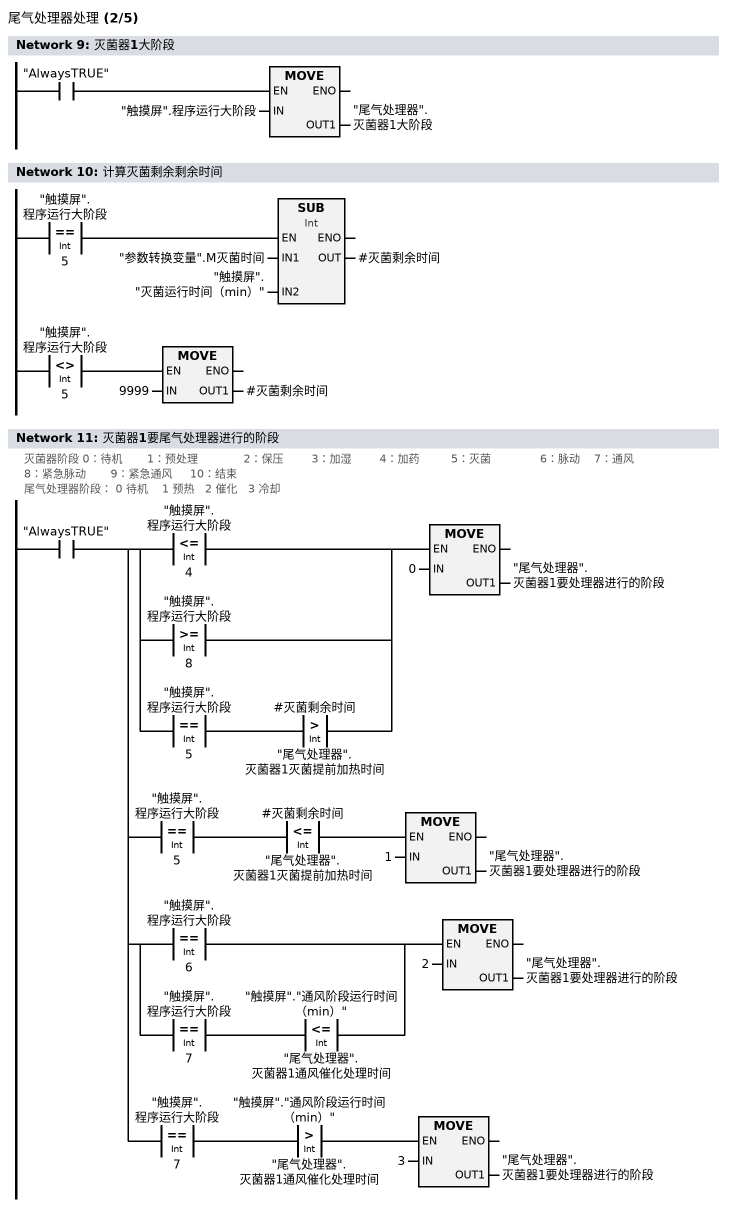
   RUNG wire#powerrail
      Contact( "AlwaysTRUE" )
      Move(in := "触摸屏".程序运行大阶段, out1 => "尾气处理器".灭菌器1大阶段)
   END_RUNG
   // the same network as SCL:
   IF "AlwaysTRUE" THEN "尾气处理器".灭菌器1大阶段 := "触摸屏".程序运行大阶段; END_IF;
END_REGION

REGION Network 10: 计算灭菌剩余剩余时间
   RUNG wire#powerrail
      { S7_Templates := "SrcType := Int" } EQ_Contact(in1 := "触摸屏".程序运行大阶段, in2 := 5)
      { S7_Templates := "SrcType := Int" } Sub(in1 := "参数转换变量".M灭菌时间, in2 := "触摸屏"."灭菌运行时间（min）", out => #灭菌剩余时间)
   END_RUNG
   RUNG wire#powerrail
      { S7_Templates := "SrcType := Int" } NE_Contact(in1 := "触摸屏".程序运行大阶段, in2 := 5)
      Move(in := 9999, out1 => #灭菌剩余时间)
   END_RUNG
   // the same network as SCL:
   IF "触摸屏".程序运行大阶段 = 5 THEN #灭菌剩余时间 := "参数转换变量".M灭菌时间 - "触摸屏"."灭菌运行时间（min）"; END_IF;
   IF "触摸屏".程序运行大阶段 <> 5 THEN #灭菌剩余时间 := 9999; END_IF;
END_REGION

REGION Network 11: 灭菌器1要尾气处理器进行的阶段
   // 灭菌器阶段 0：待机       1：预处理             2：保压        3：加湿        4：加药         5：灭菌              6：脉动    7：通风         8：紧急脉动       9：紧急通风     10：结束
   // 
   // 尾气处理器阶段： 0 待机    1 预热   2 催化   3 冷却
   RUNG wire#powerrail
      Contact( "AlwaysTRUE" )
      wire#w1
      { S7_Templates := "SrcType := Int" } LE_Contact(in1 := "触摸屏".程序运行大阶段, in2 := 4)
      wire#w2
      Move(in := 0, out1 => "尾气处理器".灭菌器1要处理器进行的阶段)
   END_RUNG
   RUNG wire#w1
      { S7_Templates := "SrcType := Int" } GE_Contact(in1 := "触摸屏".程序运行大阶段, in2 := 8)
   END_RUNG wire#w2
   RUNG wire#w1
      { S7_Templates := "SrcType := Int" } EQ_Contact(in1 := "触摸屏".程序运行大阶段, in2 := 5)
      { S7_Templates := "SrcType := Int" } GT_Contact(in1 := #灭菌剩余时间, in2 := "尾气处理器".灭菌器1灭菌提前加热时间)
   END_RUNG wire#w2
   RUNG wire#w1
      { S7_Templates := "SrcType := Int" } EQ_Contact(in1 := "触摸屏".程序运行大阶段, in2 := 5)
      { S7_Templates := "SrcType := Int" } LE_Contact(in1 := #灭菌剩余时间, in2 := "尾气处理器".灭菌器1灭菌提前加热时间)
      Move(in := 1, out1 => "尾气处理器".灭菌器1要处理器进行的阶段)
   END_RUNG
   RUNG wire#w1
      { S7_Templates := "SrcType := Int" } EQ_Contact(in1 := "触摸屏".程序运行大阶段, in2 := 6)
      wire#w3
      Move(in := 2, out1 => "尾气处理器".灭菌器1要处理器进行的阶段)
   END_RUNG
   RUNG wire#w1
      { S7_Templates := "SrcType := Int" } EQ_Contact(in1 := "触摸屏".程序运行大阶段, in2 := 7)
      { S7_Templates := "SrcType := Int" } LE_Contact(in1 := "触摸屏"."通风阶段运行时间（min）", in2 := "尾气处理器".灭菌器1通风催化处理时间)
   END_RUNG wire#w3
   RUNG wire#w1
      { S7_Templates := "SrcType := Int" } EQ_Contact(in1 := "触摸屏".程序运行大阶段, in2 := 7)
      { S7_Templates := "SrcType := Int" } GT_Contact(in1 := "触摸屏"."通风阶段运行时间（min）", in2 := "尾气处理器".灭菌器1通风催化处理时间)
      Move(in := 3, out1 => "尾气处理器".灭菌器1要处理器进行的阶段)
   END_RUNG
   // the same network as SCL:
   IF "AlwaysTRUE" AND (("触摸屏".程序运行大阶段 <= 4) OR ("触摸屏".程序运行大阶段 >= 8) OR (("触摸屏".程序运行大阶段 = 5) AND (#灭菌剩余时间 > "尾气处理器".灭菌器1灭菌提前加热时间))) THEN
       "尾气处理器".灭菌器1要处理器进行的阶段 := 0;
   END_IF;
   IF "AlwaysTRUE" AND ("触摸屏".程序运行大阶段 = 5) AND (#灭菌剩余时间 <= "尾气处理器".灭菌器1灭菌提前加热时间) THEN
       "尾气处理器".灭菌器1要处理器进行的阶段 := 1;
   END_IF;
   IF "AlwaysTRUE" AND (("触摸屏".程序运行大阶段 = 6) OR (("触摸屏".程序运行大阶段 = 7) AND ("触摸屏"."通风阶段运行时间（min）" <= "尾气处理器".灭菌器1通风催化处理时间))) THEN
       "尾气处理器".灭菌器1要处理器进行的阶段 := 2;
   END_IF;
   IF "AlwaysTRUE" AND ("触摸屏".程序运行大阶段 = 7) AND ("触摸屏"."通风阶段运行时间（min）" > "尾气处理器".灭菌器1通风催化处理时间) THEN
       "尾气处理器".灭菌器1要处理器进行的阶段 := 3;
   END_IF;
END_REGION

REGION Network 12: 灭菌工艺参数初始化
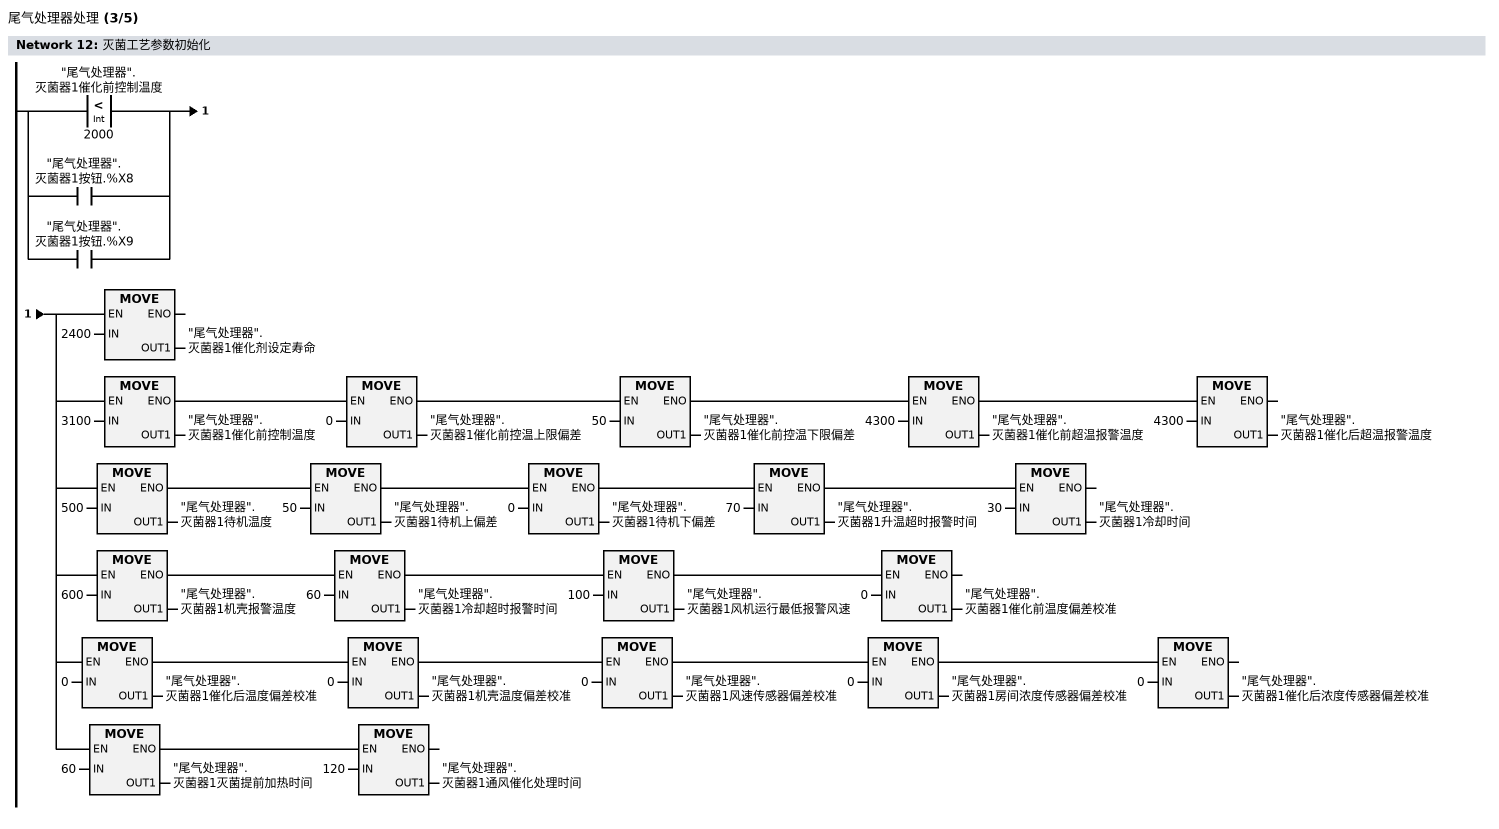
   RUNG wire#powerrail
      { S7_Templates := "SrcType := Int" } LT_Contact(in1 := "尾气处理器".灭菌器1催化前控制温度, in2 := 2000)
      wire#w1
      Move(in := 2400, out1 => "尾气处理器".灭菌器1催化剂设定寿命)
   END_RUNG
   RUNG wire#powerrail
      Contact( "尾气处理器".灭菌器1按钮.%X8 )
   END_RUNG wire#w1
   RUNG wire#powerrail
      Contact( "尾气处理器".灭菌器1按钮.%X9 )
   END_RUNG wire#w1
   RUNG wire#w1
      Move(in := 3100, out1 => "尾气处理器".灭菌器1催化前控制温度)
      Move(in := 0, out1 => "尾气处理器".灭菌器1催化前控温上限偏差)
      Move(in := 50, out1 => "尾气处理器".灭菌器1催化前控温下限偏差)
      Move(in := 4300, out1 => "尾气处理器".灭菌器1催化前超温报警温度)
      Move(in := 4300, out1 => "尾气处理器".灭菌器1催化后超温报警温度)
   END_RUNG
   RUNG wire#w1
      Move(in := 500, out1 => "尾气处理器".灭菌器1待机温度)
      Move(in := 50, out1 => "尾气处理器".灭菌器1待机上偏差)
      Move(in := 0, out1 => "尾气处理器".灭菌器1待机下偏差)
      Move(in := 70, out1 => "尾气处理器".灭菌器1升温超时报警时间)
      Move(in := 30, out1 => "尾气处理器".灭菌器1冷却时间)
   END_RUNG
   RUNG wire#w1
      Move(in := 600, out1 => "尾气处理器".灭菌器1机壳报警温度)
      Move(in := 60, out1 => "尾气处理器".灭菌器1冷却超时报警时间)
      Move(in := 100, out1 => "尾气处理器".灭菌器1风机运行最低报警风速)
      Move(in := 0, out1 => "尾气处理器".灭菌器1催化前温度偏差校准)
   END_RUNG
   RUNG wire#w1
      Move(in := 0, out1 => "尾气处理器".灭菌器1催化后温度偏差校准)
      Move(in := 0, out1 => "尾气处理器".灭菌器1机壳温度偏差校准)
      Move(in := 0, out1 => "尾气处理器".灭菌器1风速传感器偏差校准)
      Move(in := 0, out1 => "尾气处理器".灭菌器1房间浓度传感器偏差校准)
      Move(in := 0, out1 => "尾气处理器".灭菌器1催化后浓度传感器偏差校准)
   END_RUNG
   RUNG wire#w1
      Move(in := 60, out1 => "尾气处理器".灭菌器1灭菌提前加热时间)
      Move(in := 120, out1 => "尾气处理器".灭菌器1通风催化处理时间)
   END_RUNG
   // the same network as SCL:
   IF ("尾气处理器".灭菌器1催化前控制温度 < 2000) OR "尾气处理器".灭菌器1按钮.%X8 OR "尾气处理器".灭菌器1按钮.%X9 THEN
       "尾气处理器".灭菌器1催化剂设定寿命 := 2400;
   END_IF;
   #_w1 := ("尾气处理器".灭菌器1催化前控制温度 < 2000) OR "尾气处理器".灭菌器1按钮.%X8 OR "尾气处理器".灭菌器1按钮.%X9;
   #_w2 := ("尾气处理器".灭菌器1催化前控制温度 < 2000) OR "尾气处理器".灭菌器1按钮.%X8 OR "尾气处理器".灭菌器1按钮.%X9;
   IF #_w2 THEN
       "尾气处理器".灭菌器1催化前控制温度 := 3100;
       "尾气处理器".灭菌器1催化前控温上限偏差 := 0;
       "尾气处理器".灭菌器1催化前控温下限偏差 := 50;
       "尾气处理器".灭菌器1催化前超温报警温度 := 4300;
       "尾气处理器".灭菌器1催化后超温报警温度 := 4300;
   END_IF;
   IF #_w1 THEN
       "尾气处理器".灭菌器1待机温度 := 500;
       "尾气处理器".灭菌器1待机上偏差 := 50;
       "尾气处理器".灭菌器1待机下偏差 := 0;
       "尾气处理器".灭菌器1升温超时报警时间 := 70;
       "尾气处理器".灭菌器1冷却时间 := 30;
       "尾气处理器".灭菌器1机壳报警温度 := 600;
       "尾气处理器".灭菌器1冷却超时报警时间 := 60;
       "尾气处理器".灭菌器1风机运行最低报警风速 := 100;
       "尾气处理器".灭菌器1催化前温度偏差校准 := 0;
       "尾气处理器".灭菌器1催化后温度偏差校准 := 0;
       "尾气处理器".灭菌器1机壳温度偏差校准 := 0;
       "尾气处理器".灭菌器1风速传感器偏差校准 := 0;
       "尾气处理器".灭菌器1房间浓度传感器偏差校准 := 0;
       "尾气处理器".灭菌器1催化后浓度传感器偏差校准 := 0;
       "尾气处理器".灭菌器1灭菌提前加热时间 := 60;
       "尾气处理器".灭菌器1通风催化处理时间 := 120;
   END_IF;
END_REGION

REGION Network 13: 灭菌器1程序工艺参数1
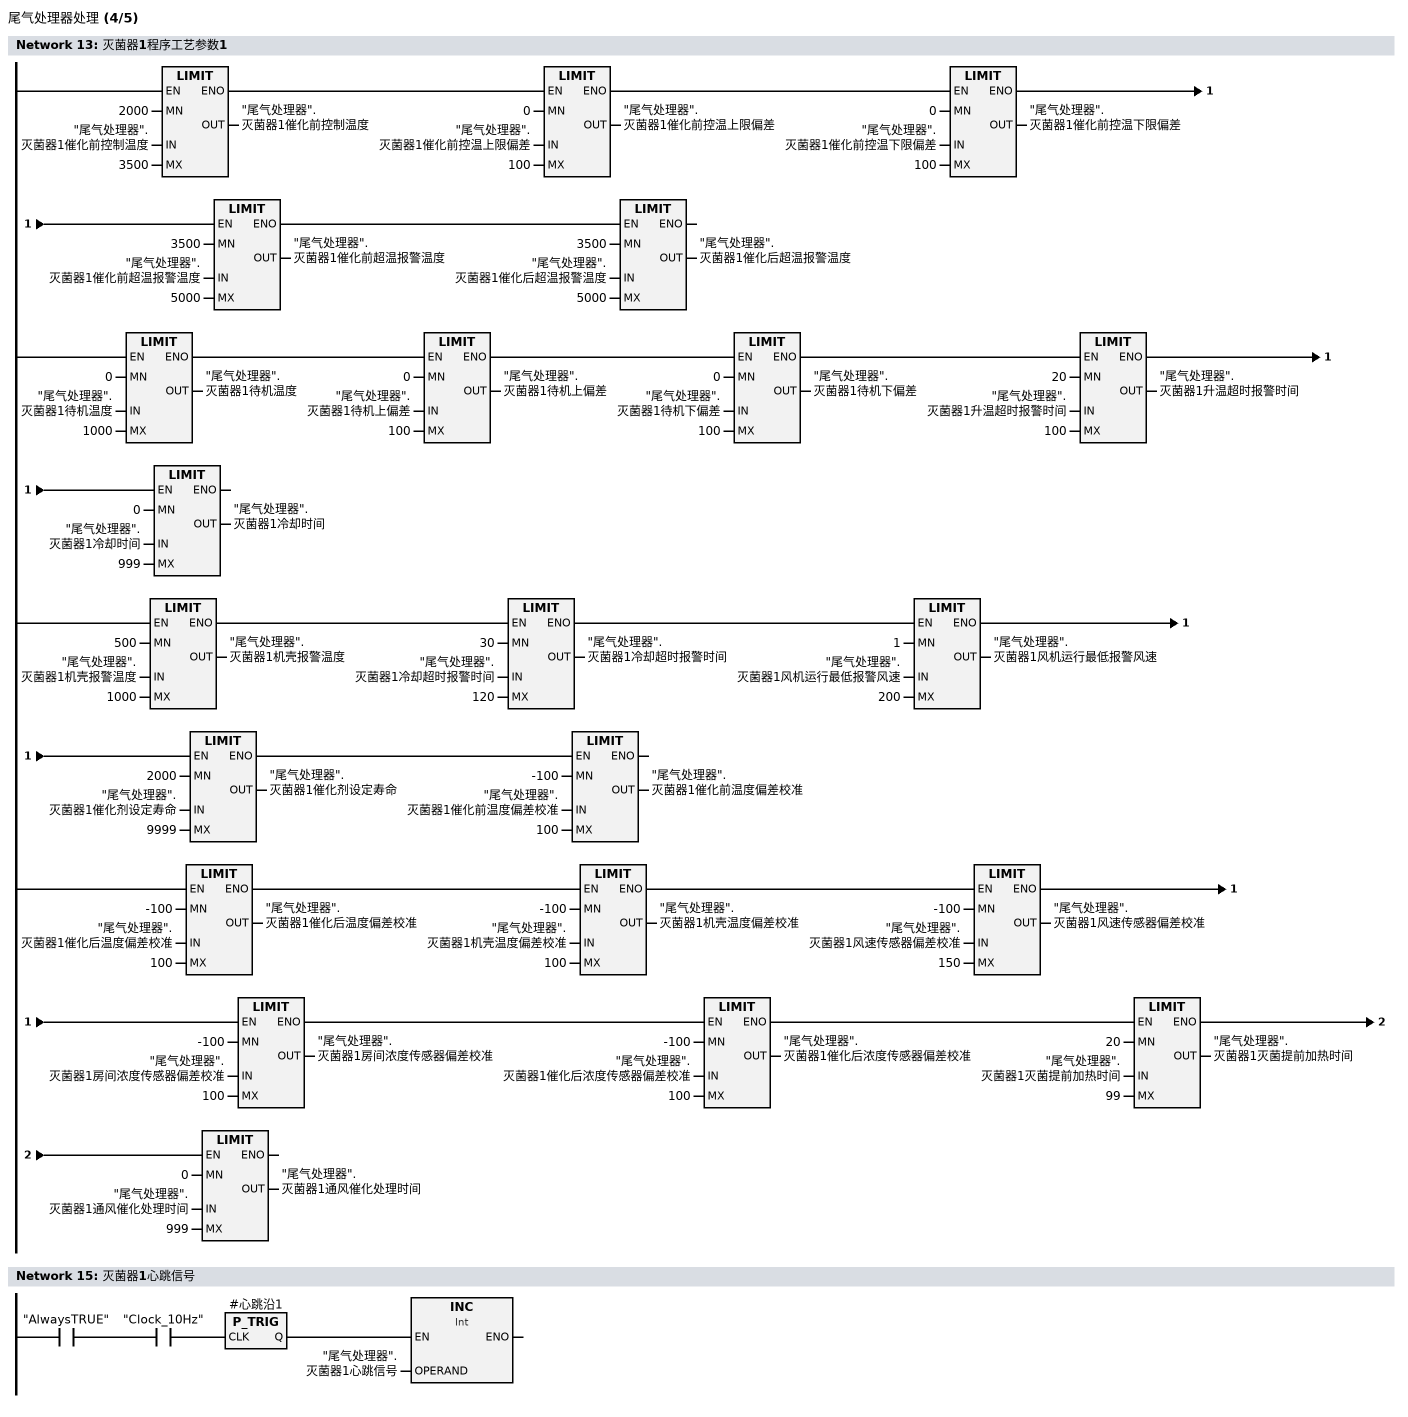
   "尾气处理器".灭菌器1催化前控制温度 := LIMIT(MN := 2000, IN := "尾气处理器".灭菌器1催化前控制温度, MX := 3500);
   "尾气处理器".灭菌器1催化前控温上限偏差 := LIMIT(MN := 0, IN := "尾气处理器".灭菌器1催化前控温上限偏差, MX := 100);
   "尾气处理器".灭菌器1催化前控温下限偏差 := LIMIT(MN := 0, IN := "尾气处理器".灭菌器1催化前控温下限偏差, MX := 100);
   "尾气处理器".灭菌器1催化前超温报警温度 := LIMIT(MN := 3500, IN := "尾气处理器".灭菌器1催化前超温报警温度, MX := 5000);
   "尾气处理器".灭菌器1催化后超温报警温度 := LIMIT(MN := 3500, IN := "尾气处理器".灭菌器1催化后超温报警温度, MX := 5000);
   "尾气处理器".灭菌器1待机温度 := LIMIT(MN := 0, IN := "尾气处理器".灭菌器1待机温度, MX := 1000);
   "尾气处理器".灭菌器1待机上偏差 := LIMIT(MN := 0, IN := "尾气处理器".灭菌器1待机上偏差, MX := 100);
   "尾气处理器".灭菌器1待机下偏差 := LIMIT(MN := 0, IN := "尾气处理器".灭菌器1待机下偏差, MX := 100);
   "尾气处理器".灭菌器1升温超时报警时间 := LIMIT(MN := 20, IN := "尾气处理器".灭菌器1升温超时报警时间, MX := 100);
   "尾气处理器".灭菌器1冷却时间 := LIMIT(MN := 0, IN := "尾气处理器".灭菌器1冷却时间, MX := 999);
   "尾气处理器".灭菌器1机壳报警温度 := LIMIT(MN := 500, IN := "尾气处理器".灭菌器1机壳报警温度, MX := 1000);
   "尾气处理器".灭菌器1冷却超时报警时间 := LIMIT(MN := 30, IN := "尾气处理器".灭菌器1冷却超时报警时间, MX := 120);
   "尾气处理器".灭菌器1风机运行最低报警风速 := LIMIT(MN := 1, IN := "尾气处理器".灭菌器1风机运行最低报警风速, MX := 200);
   "尾气处理器".灭菌器1催化剂设定寿命 := LIMIT(MN := 2000, IN := "尾气处理器".灭菌器1催化剂设定寿命, MX := 9999);
   "尾气处理器".灭菌器1催化前温度偏差校准 := LIMIT(MN := -100, IN := "尾气处理器".灭菌器1催化前温度偏差校准, MX := 100);
   "尾气处理器".灭菌器1催化后温度偏差校准 := LIMIT(MN := -100, IN := "尾气处理器".灭菌器1催化后温度偏差校准, MX := 100);
   "尾气处理器".灭菌器1机壳温度偏差校准 := LIMIT(MN := -100, IN := "尾气处理器".灭菌器1机壳温度偏差校准, MX := 100);
   "尾气处理器".灭菌器1风速传感器偏差校准 := LIMIT(MN := -100, IN := "尾气处理器".灭菌器1风速传感器偏差校准, MX := 150);
   "尾气处理器".灭菌器1房间浓度传感器偏差校准 := LIMIT(MN := -100, IN := "尾气处理器".灭菌器1房间浓度传感器偏差校准, MX := 100);
   "尾气处理器".灭菌器1催化后浓度传感器偏差校准 := LIMIT(MN := -100, IN := "尾气处理器".灭菌器1催化后浓度传感器偏差校准, MX := 100);
   "尾气处理器".灭菌器1灭菌提前加热时间 := LIMIT(MN := 20, IN := "尾气处理器".灭菌器1灭菌提前加热时间, MX := 99);
   "尾气处理器".灭菌器1通风催化处理时间 := LIMIT(MN := 0, IN := "尾气处理器".灭菌器1通风催化处理时间, MX := 999);
END_REGION

REGION Network 14: 灭菌器1程序工艺参数2
END_REGION

REGION Network 15: 灭菌器1心跳信号
   RUNG wire#powerrail
      Contact( "AlwaysTRUE" )
      Contact( "Clock_10Hz" )
      P_Trig( #心跳沿1 )
      { S7_Templates := "DestType := Int" } Inc( "尾气处理器".灭菌器1心跳信号 )
   END_RUNG
   // the same network as SCL:
   #_w1 := "AlwaysTRUE" AND "Clock_10Hz";
   #_w2 := #_w1 AND NOT #心跳沿1;   // rising edge
   #心跳沿1 := #_w1;
   IF #_w2 THEN "尾气处理器".灭菌器1心跳信号 := "尾气处理器".灭菌器1心跳信号 + 1; END_IF;
END_REGION

REGION Network 16: 灭菌器2大阶段
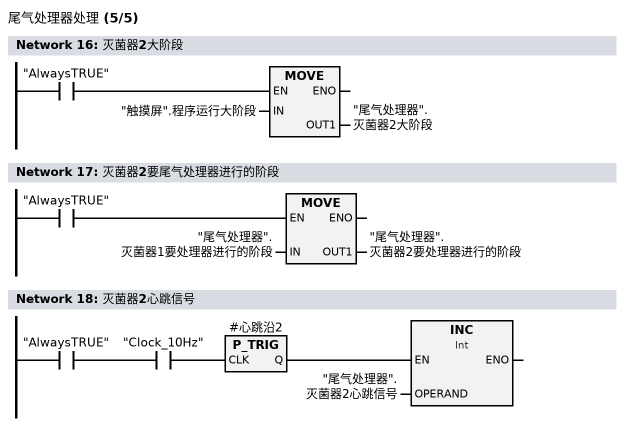
   RUNG wire#powerrail
      Contact( "AlwaysTRUE" )
      Move(in := "触摸屏".程序运行大阶段, out1 => "尾气处理器".灭菌器2大阶段)
   END_RUNG
   // the same network as SCL:
   IF "AlwaysTRUE" THEN "尾气处理器".灭菌器2大阶段 := "触摸屏".程序运行大阶段; END_IF;
END_REGION

REGION Network 17: 灭菌器2要尾气处理器进行的阶段
   RUNG wire#powerrail
      Contact( "AlwaysTRUE" )
      Move(in := "尾气处理器".灭菌器1要处理器进行的阶段, out1 => "尾气处理器".灭菌器2要处理器进行的阶段)
   END_RUNG
   // the same network as SCL:
   IF "AlwaysTRUE" THEN "尾气处理器".灭菌器2要处理器进行的阶段 := "尾气处理器".灭菌器1要处理器进行的阶段; END_IF;
END_REGION

REGION Network 18: 灭菌器2心跳信号
   RUNG wire#powerrail
      Contact( "AlwaysTRUE" )
      Contact( "Clock_10Hz" )
      P_Trig( #心跳沿2 )
      { S7_Templates := "DestType := Int" } Inc( "尾气处理器".灭菌器2心跳信号 )
   END_RUNG
   // the same network as SCL:
   #_w1 := "AlwaysTRUE" AND "Clock_10Hz";
   #_w2 := #_w1 AND NOT #心跳沿2;   // rising edge
   #心跳沿2 := #_w1;
   IF #_w2 THEN "尾气处理器".灭菌器2心跳信号 := "尾气处理器".灭菌器2心跳信号 + 1; END_IF;
END_REGION
END_FUNCTION_BLOCK

// folder: 21蜂鸣器控制

FUNCTION_BLOCK "蜂鸣器控制流程子程序"   // FB40, LAD
{ S7_Optimized_Access := 'TRUE' }
VERSION : 0.1
   VAR_INPUT
      新报警触发标志 : Bool;
      在报警画面标志 : Bool;
      报警蜂鸣器开周期 : UInt;
      报警蜂鸣器关周期 : UInt;
      报警蜂鸣器总鸣响时间 : UInt;
      在程序结束画面标志 : Bool;
      结束蜂鸣器开周期 : UInt;
      结束蜂鸣器关周期 : UInt;
      结束蜂鸣器总鸣响时间 : UInt;
   END_VAR
   VAR_OUTPUT
      蜂鸣器输出标志 : Bool;
   END_VAR
   VAR
      蜂鸣器开启时间 : UInt;
      蜂鸣器关闭时间 : UInt;
      蜂鸣器工作开关 : Bool;
      有新报警标记 : Bool;
      有新报警标记上升沿 : Bool;
      新报警时间统计沿 : Bool;
      新报警时间统计秒 : UInt;
      蜂鸣器开启时间time : Time;
      蜂鸣器关闭时间time : Time;
      有新报警并且在报警画面 : Bool;
      程序结束时间统计沿 : Bool;
      程序结束时间统计秒 : UInt;
      报警画面结束延时1s : IEC_TIMER;
      蜂鸣器开启时间ms : IEC_TIMER;
      蜂鸣器关闭时间ms : IEC_TIMER;
   END_VAR
   VAR_TEMP   // added for the SCL form of the ladder/FBD networks
      _w1 : Bool;
      _w2 : Bool;
      _w3 : Bool;
      _w4 : Bool;
      _w5 : Bool;
   END_VAR
BEGIN

REGION Network 1: 处理报警时的蜂鸣器
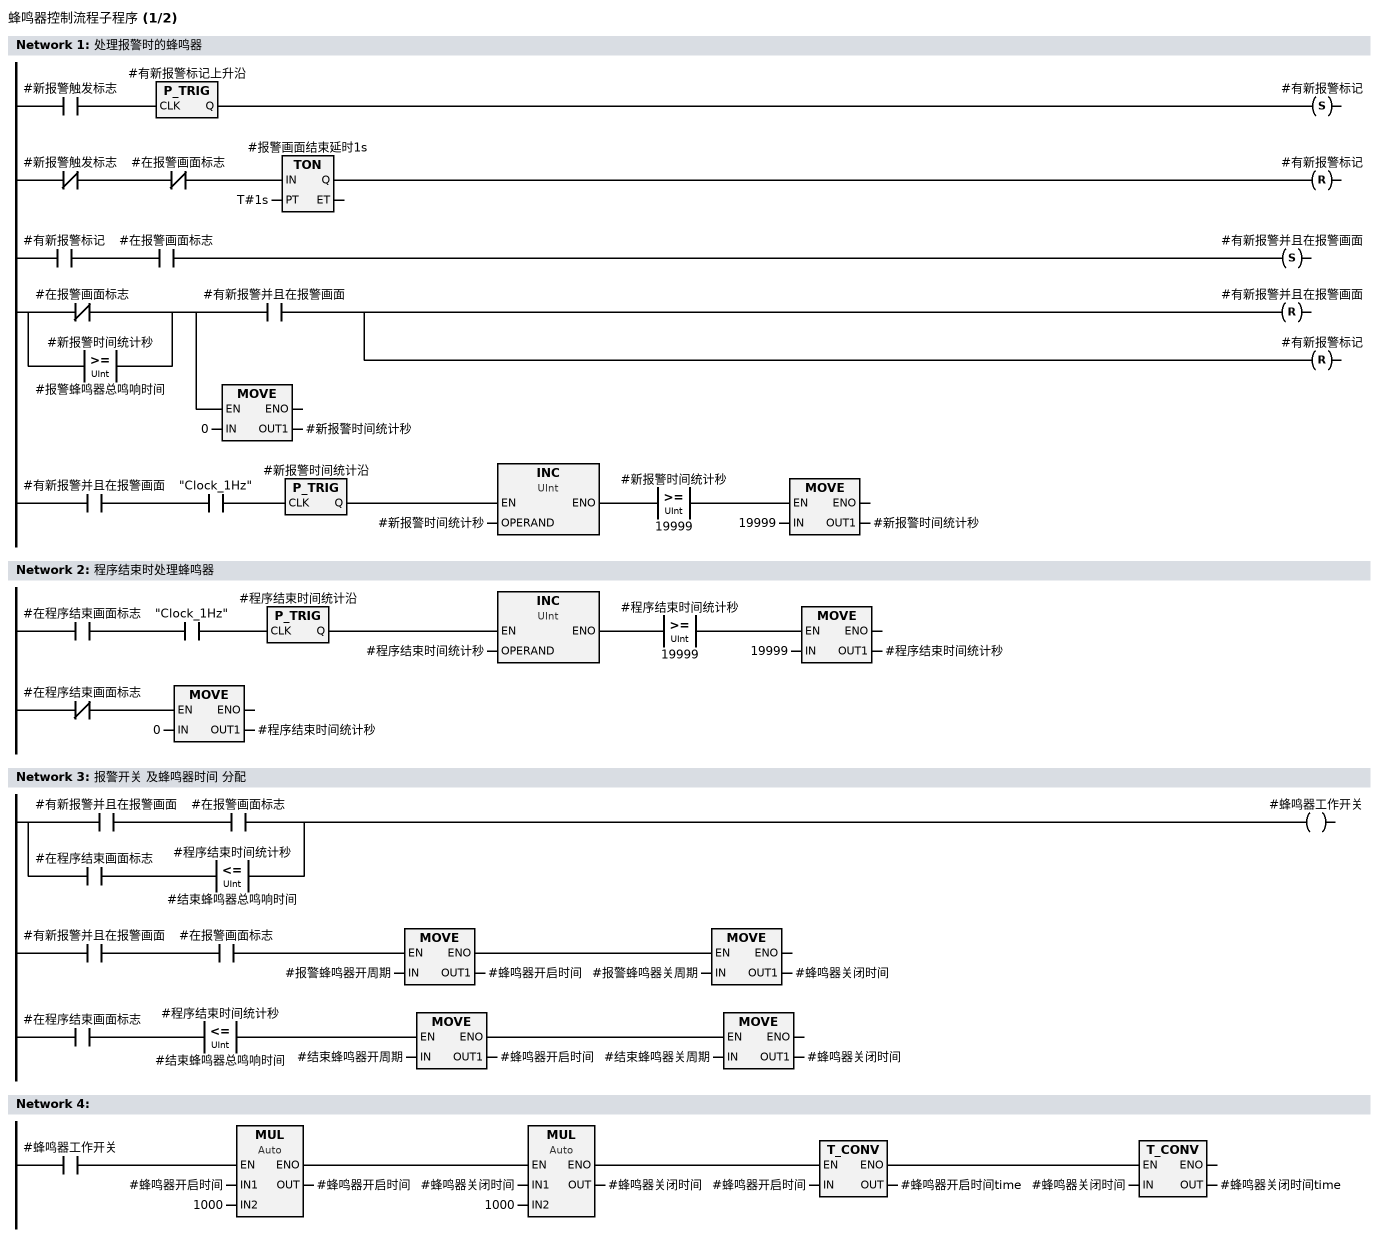
   #_w1 := #新报警触发标志 AND NOT #有新报警标记上升沿;   // rising edge
   #有新报警标记上升沿 := #新报警触发标志;
   IF #_w1 THEN #有新报警标记 := TRUE; END_IF;
   #报警画面结束延时1s.TON(IN := NOT #新报警触发标志 AND NOT #在报警画面标志, PT := T#1s);
   IF #报警画面结束延时1s.Q THEN #有新报警标记 := FALSE; END_IF;
   IF #有新报警标记 AND #在报警画面标志 THEN #有新报警并且在报警画面 := TRUE; END_IF;
   #_w2 := NOT #在报警画面标志 OR (#新报警时间统计秒 >= #报警蜂鸣器总鸣响时间);
   #_w3 := #_w2 AND #有新报警并且在报警画面;
   IF #_w3 THEN
       #有新报警并且在报警画面 := FALSE;
       #有新报警标记 := FALSE;
   END_IF;
   IF #_w2 THEN #新报警时间统计秒 := 0; END_IF;
   #_w4 := #有新报警并且在报警画面 AND "Clock_1Hz";
   #_w5 := #_w4 AND NOT #新报警时间统计沿;   // rising edge
   #新报警时间统计沿 := #_w4;
   IF #_w5 THEN #新报警时间统计秒 := #新报警时间统计秒 + 1; END_IF;
   IF #_w5 AND (#新报警时间统计秒 >= 19999) THEN #新报警时间统计秒 := 19999; END_IF;
END_REGION

REGION Network 2: 程序结束时处理蜂鸣器
   RUNG wire#powerrail
      Contact( #在程序结束画面标志 )
      Contact( "Clock_1Hz" )
      P_Trig( #程序结束时间统计沿 )
      { S7_Templates := "DestType := UInt" } Inc( #程序结束时间统计秒 )
      { S7_Templates := "SrcType := UInt" } GE_Contact(in1 := #程序结束时间统计秒, in2 := 19999)
      Move(in := 19999, out1 => #程序结束时间统计秒)
   END_RUNG
   RUNG wire#powerrail
      I_Contact( #在程序结束画面标志 )
      Move(in := 0, out1 => #程序结束时间统计秒)
   END_RUNG
   // the same network as SCL:
   #_w1 := #在程序结束画面标志 AND "Clock_1Hz";
   #_w2 := #_w1 AND NOT #程序结束时间统计沿;   // rising edge
   #程序结束时间统计沿 := #_w1;
   IF #_w2 THEN #程序结束时间统计秒 := #程序结束时间统计秒 + 1; END_IF;
   IF #_w2 AND (#程序结束时间统计秒 >= 19999) THEN #程序结束时间统计秒 := 19999; END_IF;
   IF NOT #在程序结束画面标志 THEN #程序结束时间统计秒 := 0; END_IF;
END_REGION

REGION Network 3: 报警开关 及蜂鸣器时间 分配
   RUNG wire#powerrail
      Contact( #有新报警并且在报警画面 )
      Contact( #在报警画面标志 )
      wire#w1
      Coil( #蜂鸣器工作开关 )
   END_RUNG
   RUNG wire#powerrail
      Contact( #在程序结束画面标志 )
      { S7_Templates := "SrcType := UInt" } LE_Contact(in1 := #程序结束时间统计秒, in2 := #结束蜂鸣器总鸣响时间)
   END_RUNG wire#w1
   RUNG wire#powerrail
      Contact( #有新报警并且在报警画面 )
      Contact( #在报警画面标志 )
      Move(in := #报警蜂鸣器开周期, out1 => #蜂鸣器开启时间)
      Move(in := #报警蜂鸣器关周期, out1 => #蜂鸣器关闭时间)
   END_RUNG
   RUNG wire#powerrail
      Contact( #在程序结束画面标志 )
      { S7_Templates := "SrcType := UInt" } LE_Contact(in1 := #程序结束时间统计秒, in2 := #结束蜂鸣器总鸣响时间)
      Move(in := #结束蜂鸣器开周期, out1 => #蜂鸣器开启时间)
      Move(in := #结束蜂鸣器关周期, out1 => #蜂鸣器关闭时间)
   END_RUNG
   // the same network as SCL:
   #蜂鸣器工作开关 := (#有新报警并且在报警画面 AND #在报警画面标志) OR (#在程序结束画面标志 AND (#程序结束时间统计秒 <= #结束蜂鸣器总鸣响时间));
   IF #有新报警并且在报警画面 AND #在报警画面标志 THEN
       #蜂鸣器开启时间 := #报警蜂鸣器开周期;
       #蜂鸣器关闭时间 := #报警蜂鸣器关周期;
   END_IF;
   IF #在程序结束画面标志 AND (#程序结束时间统计秒 <= #结束蜂鸣器总鸣响时间) THEN
       #蜂鸣器开启时间 := #结束蜂鸣器开周期;
       #蜂鸣器关闭时间 := #结束蜂鸣器关周期;
   END_IF;
END_REGION

REGION Network 4
   // ENO of a box is taken as its EN; it also drops when the box reports an error
   IF #蜂鸣器工作开关 THEN
       #蜂鸣器开启时间 := #蜂鸣器开启时间 * 1000;
       #蜂鸣器关闭时间 := #蜂鸣器关闭时间 * 1000;
       #蜂鸣器开启时间time := T_CONV(IN := #蜂鸣器开启时间);
       #蜂鸣器关闭时间time := T_CONV(IN := #蜂鸣器关闭时间);
   END_IF;
END_REGION

REGION Network 5: 蜂鸣器输出周期
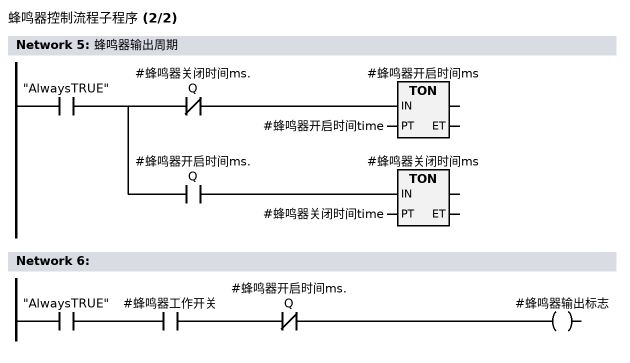
   #蜂鸣器开启时间ms.TON(IN := "AlwaysTRUE" AND NOT #蜂鸣器关闭时间ms.Q, PT := #蜂鸣器开启时间time);
   #蜂鸣器关闭时间ms.TON(IN := "AlwaysTRUE" AND #蜂鸣器开启时间ms.Q, PT := #蜂鸣器关闭时间time);
END_REGION

REGION Network 6
   RUNG wire#powerrail
      Contact( "AlwaysTRUE" )
      Contact( #蜂鸣器工作开关 )
      I_Contact( #蜂鸣器开启时间ms.Q )
      Coil( #蜂鸣器输出标志 )
   END_RUNG
   // the same network as SCL:
   #蜂鸣器输出标志 := "AlwaysTRUE" AND #蜂鸣器工作开关 AND NOT #蜂鸣器开启时间ms.Q;
END_REGION
END_FUNCTION_BLOCK

// folder: 2系统时钟

FUNCTION "系统时钟" : Void   // FC7, LAD
{ S7_Optimized_Access := 'TRUE' }
VERSION : 0.1
   VAR_INPUT
      设定年 : Int;
      设定月 : Int;
      设定日 : Int;
      设定时 : Int;
      设定分 : Int;
      设定秒 : Int;
   END_VAR
   VAR_OUTPUT
      获取年 : Int;
      获取月 : Int;
      获取日 : Int;
      获取时 : Int;
      获取分 : Int;
      获取秒 : Int;
   END_VAR
   VAR_TEMP
      获取系统时间 : DTL;
      获取系统时间完成标志 : Int;
      设定系统时间 : DTL;
      设定系统时间完成标志 : Int;
      余数 : Int;
   END_VAR
   VAR_TEMP   // added for the SCL form of the ladder/FBD networks
      _w1 : Bool;
   END_VAR
BEGIN

REGION Network 1: 读取系统时间
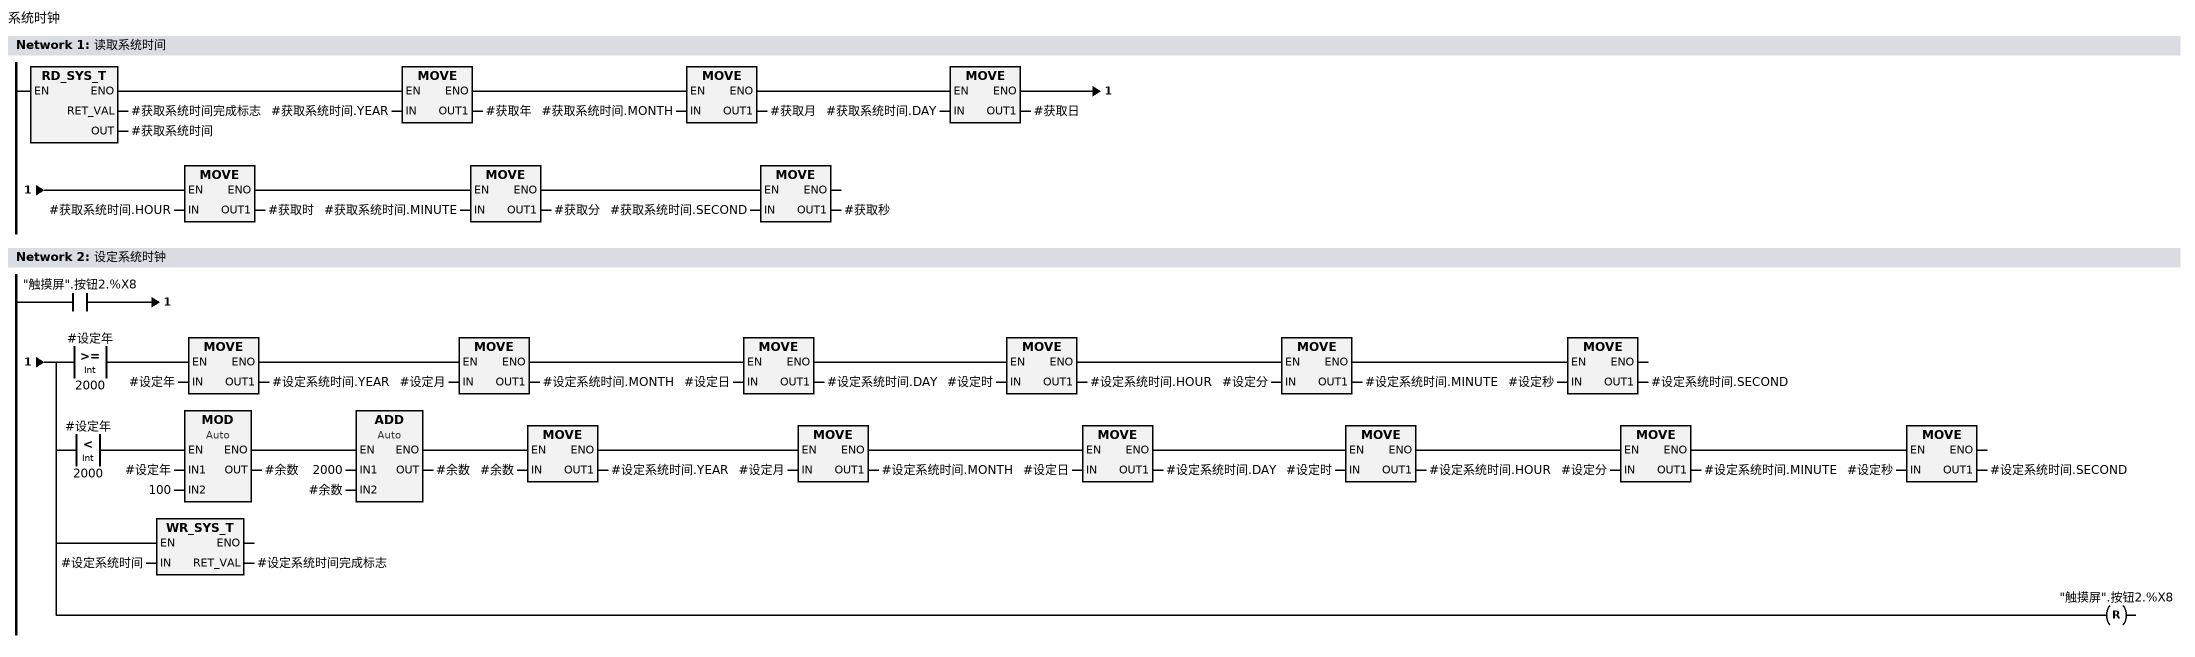
   // ENO of a box is taken as its EN; it also drops when the box reports an error
   #获取系统时间完成标志 := RD_SYS_T(OUT => #获取系统时间);
   #获取年 := #获取系统时间.YEAR;
   #获取月 := #获取系统时间.MONTH;
   #获取日 := #获取系统时间.DAY;
   #获取时 := #获取系统时间.HOUR;
   #获取分 := #获取系统时间.MINUTE;
   #获取秒 := #获取系统时间.SECOND;
END_REGION

REGION Network 2: 设定系统时钟
   IF "触摸屏".按钮2.%X8 AND (#设定年 >= 2000) THEN
       #设定系统时间.YEAR := #设定年;
       #设定系统时间.MONTH := #设定月;
       #设定系统时间.DAY := #设定日;
       #设定系统时间.HOUR := #设定时;
       #设定系统时间.MINUTE := #设定分;
       #设定系统时间.SECOND := #设定秒;
   END_IF;
   IF "触摸屏".按钮2.%X8 AND (#设定年 < 2000) THEN
       #余数 := #设定年 MOD 100;
       #余数 := 2000 + #余数;
       #设定系统时间.YEAR := #余数;
       #设定系统时间.MONTH := #设定月;
       #设定系统时间.DAY := #设定日;
       #设定系统时间.HOUR := #设定时;
       #设定系统时间.MINUTE := #设定分;
       #设定系统时间.SECOND := #设定秒;
   END_IF;
   #_w1 := "触摸屏".按钮2.%X8;
   IF #_w1 THEN
       #设定系统时间完成标志 := WR_SYS_T(IN := #设定系统时间);
       "触摸屏".按钮2.%X8 := FALSE;
   END_IF;
END_REGION
END_FUNCTION

// folder: 3报警处理

FUNCTION_BLOCK "报警处理"   // FB17, LAD
{ S7_Optimized_Access := 'TRUE' }
VERSION : 0.1
   VAR
      程序报警退出标志 : Bool;
      程序报警暂停标志 : Bool;
      程序报警脉动标志 : Bool;
      沿1 : Bool;
      抽空超时沿 : Bool;
   END_VAR
   VAR_TEMP
      小阶段名称 : Int;
   END_VAR
   VAR_TEMP   // added for the SCL form of the ladder/FBD networks
      _w1 : Bool;
      _w2 : Bool;
   END_VAR
BEGIN

REGION Network 1: A001 定期维护，请联系客服工程师
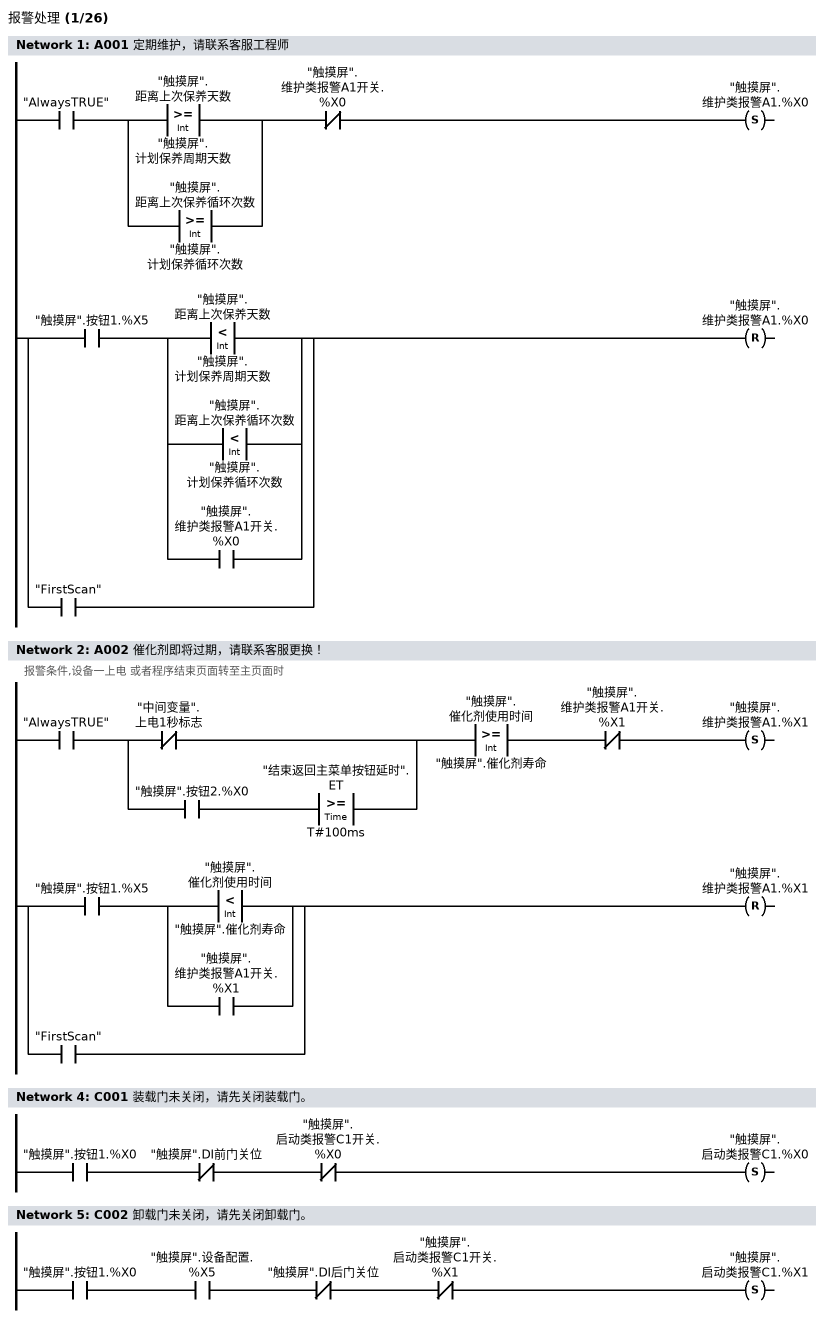
   RUNG wire#powerrail
      Contact( "AlwaysTRUE" )
      wire#w1
      { S7_Templates := "SrcType := Int" } GE_Contact(in1 := "触摸屏".距离上次保养天数, in2 := "触摸屏".计划保养周期天数)
      wire#w2
      I_Contact( "触摸屏".维护类报警A1开关.%X0 )
      S_Coil( "触摸屏".维护类报警A1.%X0 )
   END_RUNG
   RUNG wire#w1
      { S7_Templates := "SrcType := Int" } GE_Contact(in1 := "触摸屏".距离上次保养循环次数, in2 := "触摸屏".计划保养循环次数)
   END_RUNG wire#w2
   RUNG wire#powerrail
      Contact( "触摸屏".按钮1.%X5 )
      wire#w3
      { S7_Templates := "SrcType := Int" } LT_Contact(in1 := "触摸屏".距离上次保养天数, in2 := "触摸屏".计划保养周期天数)
      wire#w4
      R_Coil( "触摸屏".维护类报警A1.%X0 )
   END_RUNG
   RUNG wire#w3
      { S7_Templates := "SrcType := Int" } LT_Contact(in1 := "触摸屏".距离上次保养循环次数, in2 := "触摸屏".计划保养循环次数)
   END_RUNG wire#w4
   RUNG wire#w3
      Contact( "触摸屏".维护类报警A1开关.%X0 )
   END_RUNG wire#w4
   RUNG wire#powerrail
      Contact( "FirstScan" )
   END_RUNG wire#w4
   // the same network as SCL:
   IF "AlwaysTRUE" AND (("触摸屏".距离上次保养天数 >= "触摸屏".计划保养周期天数) OR ("触摸屏".距离上次保养循环次数 >= "触摸屏".计划保养循环次数)) AND NOT "触摸屏".维护类报警A1开关.%X0 THEN
       "触摸屏".维护类报警A1.%X0 := TRUE;
   END_IF;
   IF ("触摸屏".按钮1.%X5 AND (("触摸屏".距离上次保养天数 < "触摸屏".计划保养周期天数) OR ("触摸屏".距离上次保养循环次数 < "触摸屏".计划保养循环次数) OR "触摸屏".维护类报警A1开关.%X0)) OR "FirstScan" THEN
       "触摸屏".维护类报警A1.%X0 := FALSE;
   END_IF;
END_REGION

REGION Network 2: A002 催化剂即将过期，请联系客服更换！
   // 报警条件,设备一上电 或者程序结束页面转至主页面时
   RUNG wire#powerrail
      Contact( "AlwaysTRUE" )
      wire#w1
      I_Contact( "中间变量".上电1秒标志 )
      wire#w2
      { S7_Templates := "SrcType := Int" } GE_Contact(in1 := "触摸屏".催化剂使用时间, in2 := "触摸屏".催化剂寿命)
      I_Contact( "触摸屏".维护类报警A1开关.%X1 )
      S_Coil( "触摸屏".维护类报警A1.%X1 )
   END_RUNG
   RUNG wire#w1
      Contact( "触摸屏".按钮2.%X0 )
      { S7_Templates := "SrcType := Time" } GE_Contact(in1 := "结束返回主菜单按钮延时".ET, in2 := T#100ms)
   END_RUNG wire#w2
   RUNG wire#powerrail
      Contact( "触摸屏".按钮1.%X5 )
      wire#w3
      { S7_Templates := "SrcType := Int" } LT_Contact(in1 := "触摸屏".催化剂使用时间, in2 := "触摸屏".催化剂寿命)
      wire#w4
      R_Coil( "触摸屏".维护类报警A1.%X1 )
   END_RUNG
   RUNG wire#w3
      Contact( "触摸屏".维护类报警A1开关.%X1 )
   END_RUNG wire#w4
   RUNG wire#powerrail
      Contact( "FirstScan" )
   END_RUNG wire#w4
   // the same network as SCL:
   IF "AlwaysTRUE" AND (NOT "中间变量".上电1秒标志 OR ("触摸屏".按钮2.%X0 AND ("结束返回主菜单按钮延时".ET >= T#100ms))) AND ("触摸屏".催化剂使用时间 >= "触摸屏".催化剂寿命) AND NOT "触摸屏".维护类报警A1开关.%X1 THEN
       "触摸屏".维护类报警A1.%X1 := TRUE;
   END_IF;
   IF ("触摸屏".按钮1.%X5 AND (("触摸屏".催化剂使用时间 < "触摸屏".催化剂寿命) OR "触摸屏".维护类报警A1开关.%X1)) OR "FirstScan" THEN
       "触摸屏".维护类报警A1.%X1 := FALSE;
   END_IF;
END_REGION

REGION Network 3: 门机构相关报警B
END_REGION

REGION Network 4: C001 装载门未关闭，请先关闭装载门。
   RUNG wire#powerrail
      Contact( "触摸屏".按钮1.%X0 )
      I_Contact( "触摸屏".DI前门关位 )
      I_Contact( "触摸屏".启动类报警C1开关.%X0 )
      S_Coil( "触摸屏".启动类报警C1.%X0 )
   END_RUNG
   // the same network as SCL:
   IF "触摸屏".按钮1.%X0 AND NOT "触摸屏".DI前门关位 AND NOT "触摸屏".启动类报警C1开关.%X0 THEN "触摸屏".启动类报警C1.%X0 := TRUE; END_IF;
END_REGION

REGION Network 5: C002 卸载门未关闭，请先关闭卸载门。
   RUNG wire#powerrail
      Contact( "触摸屏".按钮1.%X0 )
      Contact( "触摸屏".设备配置.%X5 )
      I_Contact( "触摸屏".DI后门关位 )
      I_Contact( "触摸屏".启动类报警C1开关.%X1 )
      S_Coil( "触摸屏".启动类报警C1.%X1 )
   END_RUNG
   // the same network as SCL:
   IF "触摸屏".按钮1.%X0 AND "触摸屏".设备配置.%X5 AND NOT "触摸屏".DI后门关位 AND NOT "触摸屏".启动类报警C1开关.%X1 THEN
       "触摸屏".启动类报警C1.%X1 := TRUE;
   END_IF;
END_REGION

REGION Network 6: C003 内室温度过低，请等待。
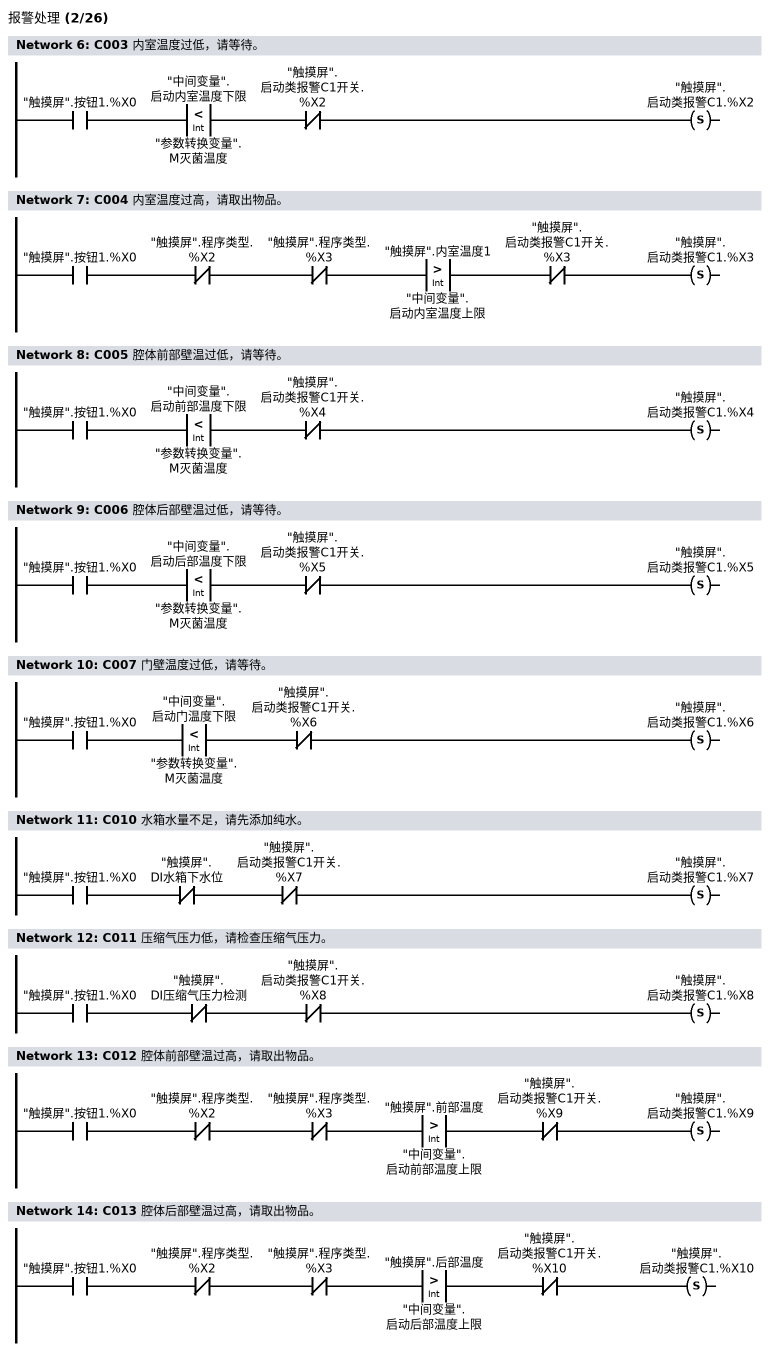
   RUNG wire#powerrail
      Contact( "触摸屏".按钮1.%X0 )
      { S7_Templates := "SrcType := Int" } LT_Contact(in1 := "中间变量".启动内室温度下限, in2 := "参数转换变量".M灭菌温度)
      I_Contact( "触摸屏".启动类报警C1开关.%X2 )
      S_Coil( "触摸屏".启动类报警C1.%X2 )
   END_RUNG
   // the same network as SCL:
   IF "触摸屏".按钮1.%X0 AND ("中间变量".启动内室温度下限 < "参数转换变量".M灭菌温度) AND NOT "触摸屏".启动类报警C1开关.%X2 THEN
       "触摸屏".启动类报警C1.%X2 := TRUE;
   END_IF;
END_REGION

REGION Network 7: C004 内室温度过高，请取出物品。
   RUNG wire#powerrail
      Contact( "触摸屏".按钮1.%X0 )
      I_Contact( "触摸屏".程序类型.%X2 )
      I_Contact( "触摸屏".程序类型.%X3 )
      { S7_Templates := "SrcType := Int" } GT_Contact(in1 := "触摸屏".内室温度1, in2 := "中间变量".启动内室温度上限)
      I_Contact( "触摸屏".启动类报警C1开关.%X3 )
      S_Coil( "触摸屏".启动类报警C1.%X3 )
   END_RUNG
   // the same network as SCL:
   IF "触摸屏".按钮1.%X0 AND NOT "触摸屏".程序类型.%X2 AND NOT "触摸屏".程序类型.%X3 AND ("触摸屏".内室温度1 > "中间变量".启动内室温度上限) AND NOT "触摸屏".启动类报警C1开关.%X3 THEN
       "触摸屏".启动类报警C1.%X3 := TRUE;
   END_IF;
END_REGION

REGION Network 8: C005 腔体前部壁温过低，请等待。
   RUNG wire#powerrail
      Contact( "触摸屏".按钮1.%X0 )
      { S7_Templates := "SrcType := Int" } LT_Contact(in1 := "中间变量".启动前部温度下限, in2 := "参数转换变量".M灭菌温度)
      I_Contact( "触摸屏".启动类报警C1开关.%X4 )
      S_Coil( "触摸屏".启动类报警C1.%X4 )
   END_RUNG
   // the same network as SCL:
   IF "触摸屏".按钮1.%X0 AND ("中间变量".启动前部温度下限 < "参数转换变量".M灭菌温度) AND NOT "触摸屏".启动类报警C1开关.%X4 THEN
       "触摸屏".启动类报警C1.%X4 := TRUE;
   END_IF;
END_REGION

REGION Network 9: C006 腔体后部壁温过低，请等待。
   RUNG wire#powerrail
      Contact( "触摸屏".按钮1.%X0 )
      { S7_Templates := "SrcType := Int" } LT_Contact(in1 := "中间变量".启动后部温度下限, in2 := "参数转换变量".M灭菌温度)
      I_Contact( "触摸屏".启动类报警C1开关.%X5 )
      S_Coil( "触摸屏".启动类报警C1.%X5 )
   END_RUNG
   // the same network as SCL:
   IF "触摸屏".按钮1.%X0 AND ("中间变量".启动后部温度下限 < "参数转换变量".M灭菌温度) AND NOT "触摸屏".启动类报警C1开关.%X5 THEN
       "触摸屏".启动类报警C1.%X5 := TRUE;
   END_IF;
END_REGION

REGION Network 10: C007 门壁温度过低，请等待。
   RUNG wire#powerrail
      Contact( "触摸屏".按钮1.%X0 )
      { S7_Templates := "SrcType := Int" } LT_Contact(in1 := "中间变量".启动门温度下限, in2 := "参数转换变量".M灭菌温度)
      I_Contact( "触摸屏".启动类报警C1开关.%X6 )
      S_Coil( "触摸屏".启动类报警C1.%X6 )
   END_RUNG
   // the same network as SCL:
   IF "触摸屏".按钮1.%X0 AND ("中间变量".启动门温度下限 < "参数转换变量".M灭菌温度) AND NOT "触摸屏".启动类报警C1开关.%X6 THEN
       "触摸屏".启动类报警C1.%X6 := TRUE;
   END_IF;
END_REGION

REGION Network 11: C010 水箱水量不足，请先添加纯水。
   RUNG wire#powerrail
      Contact( "触摸屏".按钮1.%X0 )
      I_Contact( "触摸屏".DI水箱下水位 )
      I_Contact( "触摸屏".启动类报警C1开关.%X7 )
      S_Coil( "触摸屏".启动类报警C1.%X7 )
   END_RUNG
   // the same network as SCL:
   IF "触摸屏".按钮1.%X0 AND NOT "触摸屏".DI水箱下水位 AND NOT "触摸屏".启动类报警C1开关.%X7 THEN "触摸屏".启动类报警C1.%X7 := TRUE; END_IF;
END_REGION

REGION Network 12: C011 压缩气压力低，请检查压缩气压力。
   RUNG wire#powerrail
      Contact( "触摸屏".按钮1.%X0 )
      I_Contact( "触摸屏".DI压缩气压力检测 )
      I_Contact( "触摸屏".启动类报警C1开关.%X8 )
      S_Coil( "触摸屏".启动类报警C1.%X8 )
   END_RUNG
   // the same network as SCL:
   IF "触摸屏".按钮1.%X0 AND NOT "触摸屏".DI压缩气压力检测 AND NOT "触摸屏".启动类报警C1开关.%X8 THEN
       "触摸屏".启动类报警C1.%X8 := TRUE;
   END_IF;
END_REGION

REGION Network 13: C012 腔体前部壁温过高，请取出物品。
   RUNG wire#powerrail
      Contact( "触摸屏".按钮1.%X0 )
      I_Contact( "触摸屏".程序类型.%X2 )
      I_Contact( "触摸屏".程序类型.%X3 )
      { S7_Templates := "SrcType := Int" } GT_Contact(in1 := "触摸屏".前部温度, in2 := "中间变量".启动前部温度上限)
      I_Contact( "触摸屏".启动类报警C1开关.%X9 )
      S_Coil( "触摸屏".启动类报警C1.%X9 )
   END_RUNG
   // the same network as SCL:
   IF "触摸屏".按钮1.%X0 AND NOT "触摸屏".程序类型.%X2 AND NOT "触摸屏".程序类型.%X3 AND ("触摸屏".前部温度 > "中间变量".启动前部温度上限) AND NOT "触摸屏".启动类报警C1开关.%X9 THEN
       "触摸屏".启动类报警C1.%X9 := TRUE;
   END_IF;
END_REGION

REGION Network 14: C013 腔体后部壁温过高，请取出物品。
   RUNG wire#powerrail
      Contact( "触摸屏".按钮1.%X0 )
      I_Contact( "触摸屏".程序类型.%X2 )
      I_Contact( "触摸屏".程序类型.%X3 )
      { S7_Templates := "SrcType := Int" } GT_Contact(in1 := "触摸屏".后部温度, in2 := "中间变量".启动后部温度上限)
      I_Contact( "触摸屏".启动类报警C1开关.%X10 )
      S_Coil( "触摸屏".启动类报警C1.%X10 )
   END_RUNG
   // the same network as SCL:
   IF "触摸屏".按钮1.%X0 AND NOT "触摸屏".程序类型.%X2 AND NOT "触摸屏".程序类型.%X3 AND ("触摸屏".后部温度 > "中间变量".启动后部温度上限) AND NOT "触摸屏".启动类报警C1开关.%X10 THEN
       "触摸屏".启动类报警C1.%X10 := TRUE;
   END_IF;
END_REGION

REGION Network 15: C014 门壁温度过高，请取出物品。
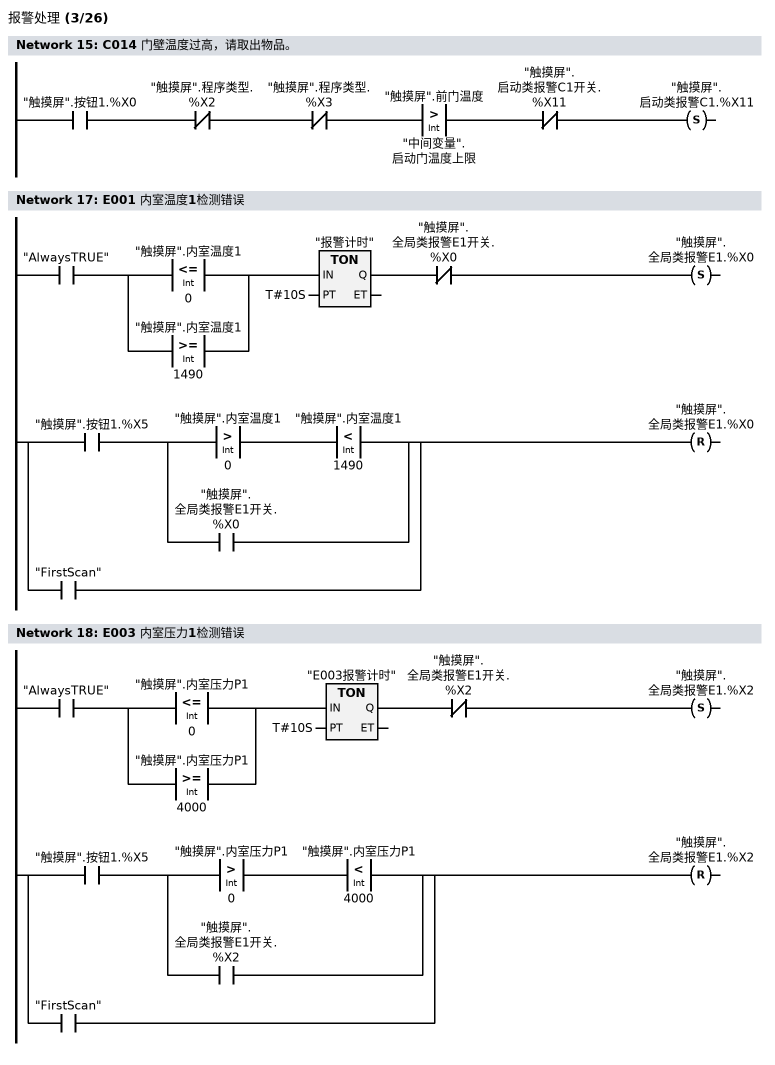
   RUNG wire#powerrail
      Contact( "触摸屏".按钮1.%X0 )
      I_Contact( "触摸屏".程序类型.%X2 )
      I_Contact( "触摸屏".程序类型.%X3 )
      { S7_Templates := "SrcType := Int" } GT_Contact(in1 := "触摸屏".前门温度, in2 := "中间变量".启动门温度上限)
      I_Contact( "触摸屏".启动类报警C1开关.%X11 )
      S_Coil( "触摸屏".启动类报警C1.%X11 )
   END_RUNG
   // the same network as SCL:
   IF "触摸屏".按钮1.%X0 AND NOT "触摸屏".程序类型.%X2 AND NOT "触摸屏".程序类型.%X3 AND ("触摸屏".前门温度 > "中间变量".启动门温度上限) AND NOT "触摸屏".启动类报警C1开关.%X11 THEN
       "触摸屏".启动类报警C1.%X11 := TRUE;
   END_IF;
END_REGION

REGION Network 16: C016 请扫描、更换气罐！
END_REGION

REGION Network 17: E001 内室温度1检测错误
   "报警计时".TON(IN := "AlwaysTRUE" AND (("触摸屏".内室温度1 <= 0) OR ("触摸屏".内室温度1 >= 1490)), PT := T#10S);
   IF "报警计时".Q AND NOT "触摸屏".全局类报警E1开关.%X0 THEN "触摸屏".全局类报警E1.%X0 := TRUE; END_IF;
   IF ("触摸屏".按钮1.%X5 AND ((("触摸屏".内室温度1 > 0) AND ("触摸屏".内室温度1 < 1490)) OR "触摸屏".全局类报警E1开关.%X0)) OR "FirstScan" THEN
       "触摸屏".全局类报警E1.%X0 := FALSE;
   END_IF;
END_REGION

REGION Network 18: E003 内室压力1检测错误
   "E003报警计时".TON(IN := "AlwaysTRUE" AND (("触摸屏".内室压力P1 <= 0) OR ("触摸屏".内室压力P1 >= 4000)), PT := T#10S);
   IF "E003报警计时".Q AND NOT "触摸屏".全局类报警E1开关.%X2 THEN "触摸屏".全局类报警E1.%X2 := TRUE; END_IF;
   IF ("触摸屏".按钮1.%X5 AND ((("触摸屏".内室压力P1 > 0) AND ("触摸屏".内室压力P1 < 4000)) OR "触摸屏".全局类报警E1开关.%X2)) OR "FirstScan" THEN
       "触摸屏".全局类报警E1.%X2 := FALSE;
   END_IF;
END_REGION

REGION Network 19: E004 内室压力2检测错误
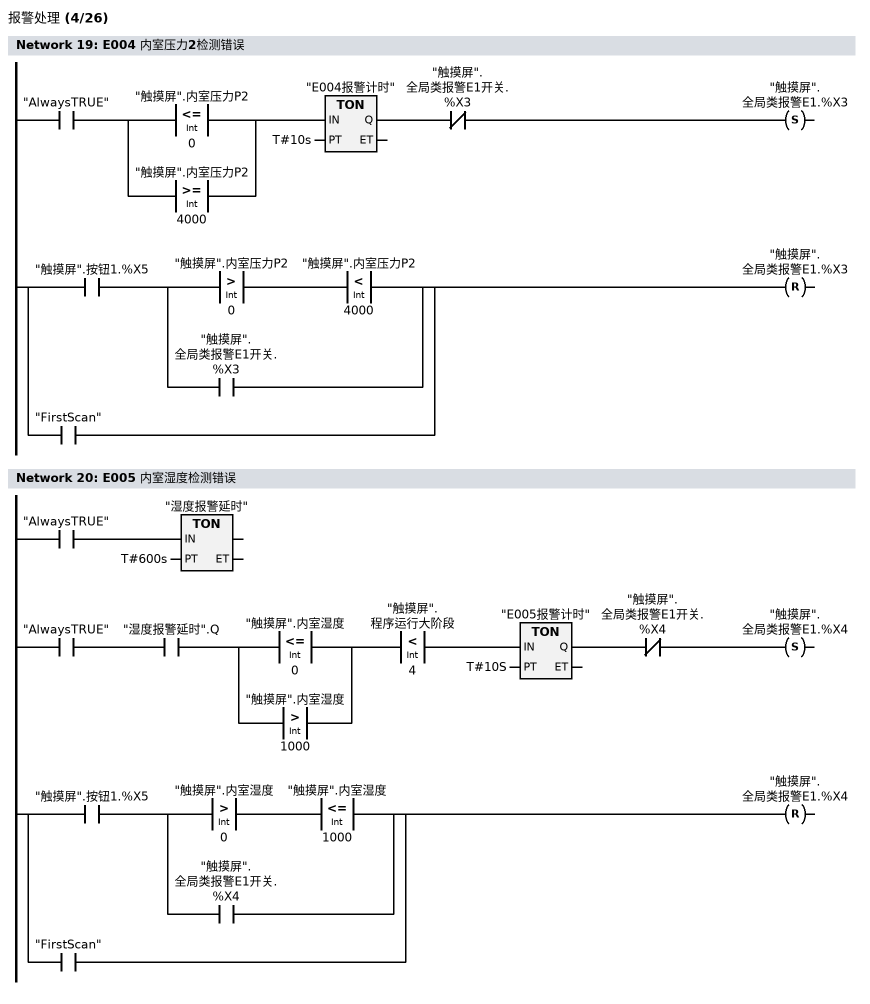
   "E004报警计时".TON(IN := "AlwaysTRUE" AND (("触摸屏".内室压力P2 <= 0) OR ("触摸屏".内室压力P2 >= 4000)), PT := T#10s);
   IF "E004报警计时".Q AND NOT "触摸屏".全局类报警E1开关.%X3 THEN "触摸屏".全局类报警E1.%X3 := TRUE; END_IF;
   IF ("触摸屏".按钮1.%X5 AND ((("触摸屏".内室压力P2 > 0) AND ("触摸屏".内室压力P2 < 4000)) OR "触摸屏".全局类报警E1开关.%X3)) OR "FirstScan" THEN
       "触摸屏".全局类报警E1.%X3 := FALSE;
   END_IF;
END_REGION

REGION Network 20: E005 内室湿度检测错误
   "湿度报警延时".TON(IN := "AlwaysTRUE", PT := T#600s);
   "E005报警计时".TON(IN := "AlwaysTRUE" AND "湿度报警延时".Q AND (("触摸屏".内室湿度 <= 0) OR ("触摸屏".内室湿度 > 1000)) AND ("触摸屏".程序运行大阶段 < 4),
                  PT := T#10S);
   IF "E005报警计时".Q AND NOT "触摸屏".全局类报警E1开关.%X4 THEN "触摸屏".全局类报警E1.%X4 := TRUE; END_IF;
   IF ("触摸屏".按钮1.%X5 AND ((("触摸屏".内室湿度 > 0) AND ("触摸屏".内室湿度 <= 1000)) OR "触摸屏".全局类报警E1开关.%X4)) OR "FirstScan" THEN
       "触摸屏".全局类报警E1.%X4 := FALSE;
   END_IF;
END_REGION

REGION Network 21: E006 腔体前部温度检测错误
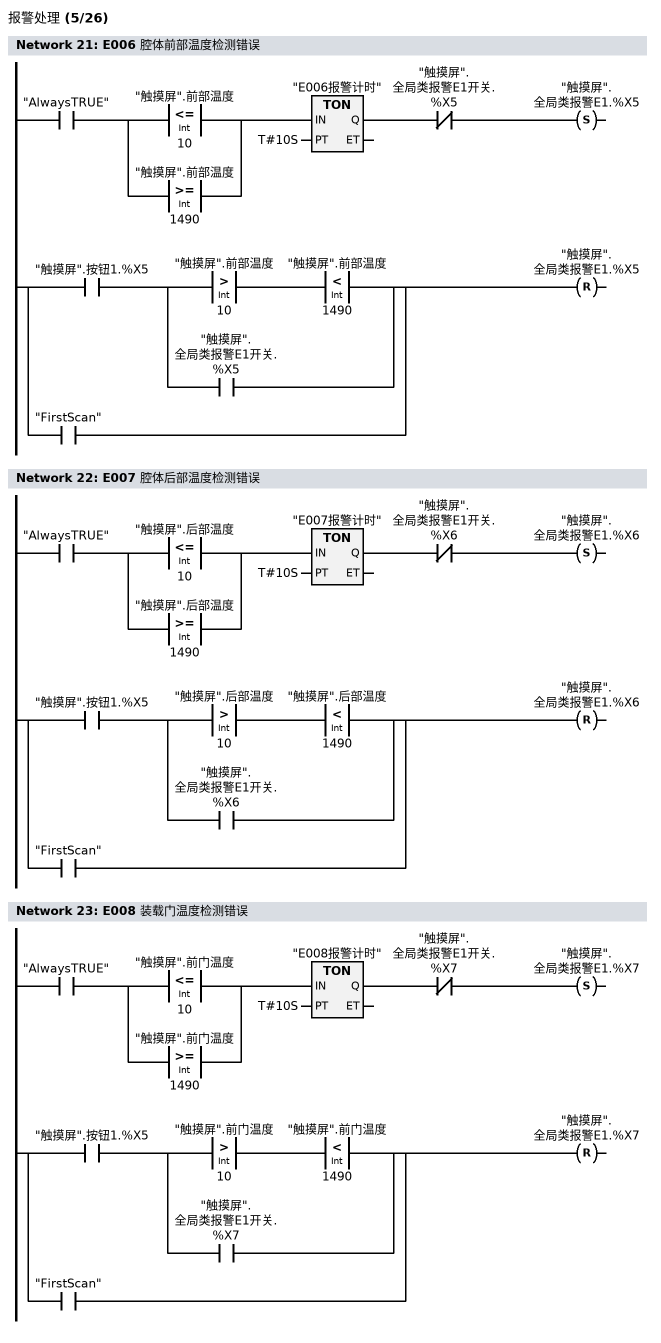
   "E006报警计时".TON(IN := "AlwaysTRUE" AND (("触摸屏".前部温度 <= 10) OR ("触摸屏".前部温度 >= 1490)), PT := T#10S);
   IF "E006报警计时".Q AND NOT "触摸屏".全局类报警E1开关.%X5 THEN "触摸屏".全局类报警E1.%X5 := TRUE; END_IF;
   IF ("触摸屏".按钮1.%X5 AND ((("触摸屏".前部温度 > 10) AND ("触摸屏".前部温度 < 1490)) OR "触摸屏".全局类报警E1开关.%X5)) OR "FirstScan" THEN
       "触摸屏".全局类报警E1.%X5 := FALSE;
   END_IF;
END_REGION

REGION Network 22: E007 腔体后部温度检测错误
   "E007报警计时".TON(IN := "AlwaysTRUE" AND (("触摸屏".后部温度 <= 10) OR ("触摸屏".后部温度 >= 1490)), PT := T#10S);
   IF "E007报警计时".Q AND NOT "触摸屏".全局类报警E1开关.%X6 THEN "触摸屏".全局类报警E1.%X6 := TRUE; END_IF;
   IF ("触摸屏".按钮1.%X5 AND ((("触摸屏".后部温度 > 10) AND ("触摸屏".后部温度 < 1490)) OR "触摸屏".全局类报警E1开关.%X6)) OR "FirstScan" THEN
       "触摸屏".全局类报警E1.%X6 := FALSE;
   END_IF;
END_REGION

REGION Network 23: E008 装载门温度检测错误
   "E008报警计时".TON(IN := "AlwaysTRUE" AND (("触摸屏".前门温度 <= 10) OR ("触摸屏".前门温度 >= 1490)), PT := T#10S);
   IF "E008报警计时".Q AND NOT "触摸屏".全局类报警E1开关.%X7 THEN "触摸屏".全局类报警E1.%X7 := TRUE; END_IF;
   IF ("触摸屏".按钮1.%X5 AND ((("触摸屏".前门温度 > 10) AND ("触摸屏".前门温度 < 1490)) OR "触摸屏".全局类报警E1开关.%X7)) OR "FirstScan" THEN
       "触摸屏".全局类报警E1.%X7 := FALSE;
   END_IF;
END_REGION

REGION Network 24: E009 汽化器温度检测错误
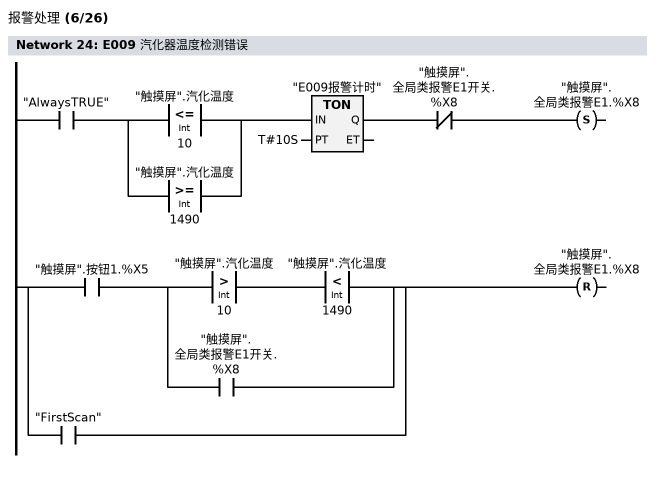
   "E009报警计时".TON(IN := "AlwaysTRUE" AND (("触摸屏".汽化温度 <= 10) OR ("触摸屏".汽化温度 >= 1490)), PT := T#10S);
   IF "E009报警计时".Q AND NOT "触摸屏".全局类报警E1开关.%X8 THEN "触摸屏".全局类报警E1.%X8 := TRUE; END_IF;
   IF ("触摸屏".按钮1.%X5 AND ((("触摸屏".汽化温度 > 10) AND ("触摸屏".汽化温度 < 1490)) OR "触摸屏".全局类报警E1开关.%X8)) OR "FirstScan" THEN
       "触摸屏".全局类报警E1.%X8 := FALSE;
   END_IF;
END_REGION

REGION Network 25: E013 加热温度过高，
   // 控制的都是前部温度的相关参数
